{region 'Documentation'}
(*!
<summary>Advances a reconciled execution slot or dispatches one first-fitting Start; no owner lifecycle changes.</summary>
*)
{endregion}
METHOD PRIVATE ProcessSlot
IF (FResult = E_Result.Error) OR FExecutionFinished THEN
    RETURN;
END_IF;
IF IsSlotCompleted() THEN
    IF IsLastSlot(Slot := FCurrentSlot) THEN
        FExecutionFinished := TRUE;
    ELSE
        SelectNextSlot();
    END_IF;
    RETURN;
END_IF;
StartNextChild();
END_METHOD

{region 'Documentation'}
(*!
<summary>Publishes technical events through the configured framework publisher.</summary>
*)
{endregion}
METHOD PRIVATE PublishEvent
VAR_INPUT
    Event : ST_Event; //! Technical event value forwarded to the selected publisher; this helper performs no retry.
END_VAR
EventPublisher.PublishEvent(Event := Event);
END_METHOD

{region 'Documentation'}
(*!
<summary>Reads one initialized child at a validated occupied index; reports invalid bindings.</summary>
*)
{endregion}
METHOD PRIVATE ReadChild : I_Orchestratable //! Initialized child interface at Index; zero on invalid access or binding, with a technical Error latched.
VAR_INPUT
    Index : DINT; //! Original array index within the cached occupied child range.
END_VAR
VAR
    Child : I_Orchestratable;
END_VAR
ReadChild := 0;
IF (FCollection = 0) OR (Index < FFirstOccupiedIndex) OR (Index > FLastOccupiedIndex) THEN
    Error(Message := CONCAT('Invalid collection access at index ', DINT_TO_STRING(Index)));
    RETURN;
END_IF;

Child := FCollection.GetChild(Index := Index);
IF Child = 0 THEN
    Error(Message := CONCAT('Missing child at index ', DINT_TO_STRING(Index)));
    RETURN;
END_IF;
IF NOT Child.IsInitialized THEN
    Error(Message := CONCAT('Uninitialized child: ', Child.Name));
    RETURN;
END_IF;

ReadChild := Child;
END_METHOD

{region 'Documentation'}
(*!
<summary>Dispatches at most one capacity-admitted Reset per call; already ready children are skipped.</summary>
*)
{endregion}
METHOD PRIVATE ResetNextChild
VAR
    Child : I_Orchestratable;
    Index : DINT;
    ReservationResult : E_EventReservationResult;
END_VAR
WHILE UDINT_TO_LINT(FNextResetOffset) < (DINT_TO_LINT(FLastOccupiedIndex) - DINT_TO_LINT(FFirstOccupiedIndex) + 1) DO
    Index := LINT_TO_DINT(DINT_TO_LINT(FFirstOccupiedIndex) + UDINT_TO_LINT(FNextResetOffset));
    Child := ReadChild(Index := Index);
    IF Child = 0 THEN
        FNextResetOffset := FNextResetOffset + 1;
        RETURN;
    END_IF;
    IF (Child.State = E_State.Idle) AND Child.IsReady THEN
        FNextResetOffset := FNextResetOffset + 1;
        CONTINUE;
    END_IF;

    ReservationResult := Child.ReserveResetEvents();
    CASE ReservationResult OF
        E_EventReservationResult.Accepted:
            Child.RequestReset();
            FNextResetOffset := FNextResetOffset + 1;
        E_EventReservationResult.WaitingForCapacity:
            RETURN;
    ELSE
        Error(Message := CONCAT('Invalid child Reset reservation: ', Child.Name));
        FNextResetOffset := FNextResetOffset + 1;
    END_CASE;
    RETURN;
END_WHILE;
END_METHOD

{region 'Documentation'}
(*!
<summary>Neutral or held technical Error; task completion is reported separately.</summary>
*)
{endregion}
{attribute 'monitoring' := 'call'}
PROPERTY PUBLIC Result : E_Result //! Neutral or held technical Error; task completion is reported separately.
GET // PUBLIC
Result := FResult;
END_GET
END_PROPERTY

{region 'Documentation'}
(*!
<summary>Selects the first or next contiguous slot group; the caller owns advancement timing.</summary>
*)
{endregion}
METHOD PRIVATE SelectNextSlot : BOOL //! TRUE after selecting a valid contiguous slot group; FALSE indicates a technical Error.
VAR
    FirstIndex : LINT;
    Slot : UDINT;
    LastIndex : DINT;
    Index : LINT;
    Child : I_Orchestratable;
    ChildSlot : UINT;
END_VAR
SelectNextSlot := FALSE;
IF FCurrentSlot = 0 THEN
    FirstIndex := DINT_TO_LINT(FFirstOccupiedIndex);
    Slot := 1;
ELSE
    FirstIndex := DINT_TO_LINT(FSlotLastIndex) + 1;
    Slot := UINT_TO_UDINT(FCurrentSlot) + 1;
END_IF;

IF (FirstIndex < DINT_TO_LINT(FFirstOccupiedIndex)) OR (FirstIndex > DINT_TO_LINT(FLastOccupiedIndex))
    OR (Slot = 0) OR (UDINT_TO_LINT(Slot) > (DINT_TO_LINT(FLastOccupiedIndex) - DINT_TO_LINT(FFirstOccupiedIndex) + 1)) THEN
    Error(Message := 'Invalid child slot boundary.');
    RETURN;
END_IF;

LastIndex := LINT_TO_DINT(FirstIndex);
FOR Index := FirstIndex TO DINT_TO_LINT(FLastOccupiedIndex) DO
    Child := ReadChild(Index := LINT_TO_DINT(Index));
    IF Child = 0 THEN
        RETURN;
    END_IF;
    ChildSlot := Child.ExecutionSlot;
    IF UINT_TO_UDINT(ChildSlot) = Slot THEN
        LastIndex := LINT_TO_DINT(Index);
        CONTINUE;
    END_IF;
    IF (Index = FirstIndex) OR (UINT_TO_UDINT(ChildSlot) <> Slot + 1) THEN
        Error(Message := 'Child slots are not contiguous and ordered.');
        RETURN;
    END_IF;
    EXIT;
END_FOR;
FCurrentSlot := UDINT_TO_UINT(Slot);
FSlotFirstIndex := LINT_TO_DINT(FirstIndex);
FSlotLastIndex := LastIndex;
SelectNextSlot := TRUE;
END_METHOD

{region 'Documentation'}
(*!
<summary>Reserves and requests at most one first-fitting Child Start within the current slot.</summary>
*)
{endregion}
METHOD PRIVATE StartNextChild
VAR
    Index : LINT;
    Child : I_Orchestratable;
    ReservationResult : E_EventReservationResult;
END_VAR
FOR Index := DINT_TO_LINT(FSlotFirstIndex) TO DINT_TO_LINT(FSlotLastIndex) DO
    Child := ReadChild(Index := LINT_TO_DINT(Index));
    IF Child = 0 THEN
        RETURN;
    END_IF;
    IF Child.State <> E_State.Idle THEN
        CONTINUE;
    END_IF;

    ReservationResult := Child.ReserveExecutionEvents();
    CASE ReservationResult OF
        E_EventReservationResult.Accepted:
            Child.RequestStart();
            FPendingStartIndex := LINT_TO_DINT(Index);
            FHasPendingStart := TRUE;
            RETURN;
        E_EventReservationResult.WaitingForCapacity:
            CONTINUE;
    ELSE
        Error(Message := CONCAT('Invalid child execution reservation: ', Child.Name));
        RETURN;
    END_CASE;
END_FOR;
END_METHOD

{region 'Documentation'}
(*!
<summary>Prepares abort completion from stopped children; no requests, diagnostics or reservation changes.</summary>
*)
{endregion}
METHOD PRIVATE UpdateAbortCompletion
VAR
    Index : LINT;
    Child : I_Orchestratable;
END_VAR
FAbortFinished := FALSE;
IF FCollection = 0 THEN
    RETURN;
END_IF;
FOR Index := DINT_TO_LINT(FFirstOccupiedIndex) TO DINT_TO_LINT(FLastOccupiedIndex) DO
    Child := FCollection.GetChild(Index := LINT_TO_DINT(Index));
    IF Child = 0 THEN
        RETURN;
    END_IF;
    IF NOT Child.IsInitialized THEN
        RETURN;
    END_IF;
    IF NOT (((Child.State = E_State.Idle) AND Child.IsReady)
        OR ((Child.State = E_State.Completed) AND Child.IsComplete)) THEN
        RETURN;
    END_IF;
END_FOR;
FAbortFinished := TRUE;
END_METHOD

{region 'Documentation'}
(*!
<summary>Prepares start readiness without interpreting previous-run results or changing children.</summary>
*)
{endregion}
METHOD PRIVATE UpdateReadiness
VAR
    Index : LINT;
    Child : I_Orchestratable;
END_VAR
FChildrenReady := FALSE;
IF FCollection = 0 THEN
    RETURN;
END_IF;
FOR Index := DINT_TO_LINT(FFirstOccupiedIndex) TO DINT_TO_LINT(FLastOccupiedIndex) DO
    Child := FCollection.GetChild(Index := LINT_TO_DINT(Index));
    IF Child = 0 THEN
        RETURN;
    END_IF;
    IF NOT Child.IsInitialized THEN
        RETURN;
    END_IF;
    IF (Child.State <> E_State.Idle) OR NOT Child.IsReady THEN
        RETURN;
    END_IF;
END_FOR;
FChildrenReady := TRUE;
END_METHOD

{region 'Documentation'}
(*!
<summary>Prepares reset completion only after all dispatch attempts; failed terminal children count as finished.</summary>
*)
{endregion}
METHOD PRIVATE UpdateResetCompletion
VAR
    Index : LINT;
    Child : I_Orchestratable;
END_VAR
FResetFinished := FALSE;
IF FCollection = 0 THEN
    RETURN;
END_IF;
IF UDINT_TO_LINT(FNextResetOffset) < (DINT_TO_LINT(FLastOccupiedIndex) - DINT_TO_LINT(FFirstOccupiedIndex) + 1) THEN
    RETURN;
END_IF;
FOR Index := DINT_TO_LINT(FFirstOccupiedIndex) TO DINT_TO_LINT(FLastOccupiedIndex) DO
    Child := FCollection.GetChild(Index := LINT_TO_DINT(Index));
    IF Child = 0 THEN
        RETURN;
    END_IF;
    IF NOT Child.IsInitialized THEN
        RETURN;
    END_IF;
    IF NOT (((Child.State = E_State.Idle) AND Child.IsReady)
        OR ((Child.State = E_State.Completed) AND Child.IsComplete)) THEN
        RETURN;
    END_IF;
END_FOR;
FResetFinished := TRUE;
END_METHOD

END_FUNCTION_BLOCK

// ---- Framework/EventBuffer/POU/FrameworkEvents/CreateFrameworkEvent.TcPOU
{region 'Documentation'}
(*!
<summary>Constructs a framework diagnostic event without publishing it.</summary>
<description>
Name and Message are ASCII text limited to the declared event capacities.
</description>
*)
{endregion}
FUNCTION CreateFrameworkEvent : ST_Event //! Constructed event value; not published. The publisher assigns SequenceId and Timestamp.
VAR_INPUT
    Name : STRING(GVL_Constants.NameLength); //! Hierarchical owner name used to identify events; must satisfy the naming contract.
    ResourceName : STRING(GVL_Constants.ResourceNameLength) := ''; //! Optional resource context for diagnostics; empty by default.
    State : E_State; //! Owner lifecycle state recorded in the event.
    Severity : E_EventSeverity; //! Logging severity for the diagnostic; independent of the test result.
    Message : STRING(GVL_Constants.MessageLength); //! Diagnostic text copied into the event within MessageLength.
END_VAR

CreateFrameworkEvent.SequenceId := 0;
CreateFrameworkEvent.Timestamp := 0;
CreateFrameworkEvent.OwnerScope := E_OwnerScope.Framework;
CreateFrameworkEvent.EventType := E_EventType.Framework;
CreateFrameworkEvent.Severity := Severity;
CreateFrameworkEvent.Name := Name;
CreateFrameworkEvent.ResourceName := ResourceName;
CreateFrameworkEvent.State := State;
CreateFrameworkEvent.Result := E_Result.NotEvaluated;
CreateFrameworkEvent.Message := Message;

END_FUNCTION

// ---- Framework/Common/POU/Stopwatch.TcPOU
{region 'Documentation'}
(*!
<summary>Internal method-driven duration measurement; no FB-body call is required. Start/Update/Stop use the current task&#x27;s scheduled timestamp. Reset clears the measurement. ElapsedTicks retains 100 ns resolution; ElapsedTime is the saturated millisecond projection.</summary>
<description>
Start replaces the previous interval. Update samples only while running and valid; Stop performs one final Update. A backward task timestamp latches invalid until Start or Reset. Property reads return held values rather than sampling the clock. ElapsedLTime is a direct conversion, without the saturation applied to ElapsedTime.


The source is the current task's scheduled timestamp, so this measures elapsed task time rather than execution cost between operations within the same task cycle. Check IsValid before using a refreshed value; a backward observation leaves the last valid duration held and does not repair itself on later Update calls.
</description>
*)
{endregion}
FUNCTION_BLOCK INTERNAL Stopwatch
VAR
    FRunning : BOOL;
    FIsValid : BOOL := TRUE;
    FStartTicks : ULINT;
    FPreviousTicks : ULINT;
    FElapsedTicks : ULINT;
END_VAR

{region 'Documentation'}
(*!
<summary>Nanosecond projection of the last updated 100 ns duration; reading does not refresh the measurement.</summary>
*)
{endregion}
{attribute 'monitoring' := 'call'}
PROPERTY PUBLIC ElapsedLTime : LTIME //! Held duration converted to LTIME nanoseconds; no refresh on read.
GET // PUBLIC
ElapsedLTime := ULINT_TO_LTIME(FElapsedTicks * 100);
END_GET
END_PROPERTY

{region 'Documentation'}
(*!
<summary>Elapsed duration in 100 ns ticks from the latest Start, Update or Stop; reading does not sample the clock.</summary>
*)
{endregion}
{attribute 'monitoring' := 'call'}
PROPERTY PUBLIC ElapsedTicks : ULINT //! Held elapsed duration in 100 ns ticks; no refresh on read.
GET // PUBLIC
ElapsedTicks := FElapsedTicks;
END_GET
END_PROPERTY

{region 'Documentation'}
(*!
<summary>Millisecond projection of the last updated duration, saturated at TIME's maximum value; reading does not refresh it.</summary>
*)
{endregion}
{attribute 'monitoring' := 'call'}
PROPERTY PUBLIC ElapsedTime : TIME //! Held duration in milliseconds, saturated at TIME's maximum; no refresh on read.
GET // PUBLIC
VAR CONSTANT
	MaxTime: ULINT := 42949672950000;
END_VAR
ElapsedTime := ULINT_TO_TIME(MIN(FElapsedTicks, MaxTime) / 10000);
END_GET
END_PROPERTY

{region 'Documentation'}
(*!
<summary>Report whether a backward clock observation has invalidated the measurement; Start or Reset restores validity.</summary>
*)
{endregion}
{attribute 'monitoring' := 'call'}
PROPERTY PUBLIC IsValid : BOOL //! FALSE after Update observes backward time; latched until Start or Reset.
GET // PUBLIC
IsValid := FIsValid;
END_GET
END_PROPERTY

{region 'Documentation'}
(*!
<summary>Clears the held measurement without starting a new interval.</summary>
*)
{endregion}
METHOD PUBLIC Reset
FRunning := FALSE;
FIsValid := TRUE;
FStartTicks := 0;
FPreviousTicks := 0;
FElapsedTicks := 0;
END_METHOD

{region 'Documentation'}
(*!
<summary>Starts a new measurement, replacing the previous value.</summary>
*)
{endregion}
METHOD PUBLIC Start
FStartTicks := Tc2_System.F_GetTaskTime();
FPreviousTicks := FStartTicks;
FElapsedTicks := 0;
FIsValid := TRUE;
FRunning := TRUE;
END_METHOD

{region 'Documentation'}
(*!
<summary>Captures the final duration and holds it until the next Start or Reset.</summary>
<description>
If the final Update detects backward time, IsValid becomes FALSE and the last valid elapsed value remains held. Stop still ends the interval. Repeated Stop calls do not sample again while stopped.
</description>
*)
{endregion}
METHOD PUBLIC Stop
Update();
FRunning := FALSE;
END_METHOD

{region 'Documentation'}
(*!
<summary>Refreshes elapsed time. A backwards clock latches invalid until Start or Reset.</summary>
*)
{endregion}
METHOD PUBLIC Update
VAR
    Ticks : ULINT;
END_VAR
IF NOT FRunning OR NOT FIsValid THEN
    RETURN;
END_IF;
Ticks := Tc2_System.F_GetTaskTime();
IF Ticks < FPreviousTicks THEN
    FIsValid := FALSE;
    RETURN;
END_IF;

FElapsedTicks := Ticks - FStartTicks;
FPreviousTicks := Ticks;
END_METHOD

END_FUNCTION_BLOCK

// ---- Framework/Common/POU/ResultAggregator.TcPOU
{region 'Documentation'}
(*!
<summary>Incrementally collect results through methods; no cyclic FB call is required. Reset starts an empty collection; Add methods always contribute. Each contribution counts once; the owner limits each collection to the UINT range.</summary>
<description>
Use Reset before each new collection and contribute each intended provider/result exactly once. AddProvider reads immediately and retains no interface. Error has highest precedence but does not stop later counter updates. TotalCount includes NotEvaluated and Abort contributions, so PassedCount, FailedCount and ErrorCount do not necessarily sum to TotalCount. The caller keeps a collection within 65535 contributions; counters are not saturating. This object emits no events and does not execute providers.
</description>
*)
{endregion}
FUNCTION_BLOCK ResultAggregator IMPLEMENTS I_ResultAggregator
VAR
    FResult : E_Result := E_Result.NotEvaluated;
    FTotalCount : UINT;
    FPassedCount : UINT;
    FFailedCount : UINT;
    FErrorCount : UINT;
END_VAR

{region 'Documentation'}
(*!
<summary>Adds one provider result; a null provider contributes one Error. Reads the result immediately; no reference is retained.</summary>
*)
{endregion}
METHOD PUBLIC AddProvider
VAR_INPUT
    Provider : I_ResultProvider; //! Result provider read immediately; zero contributes Error. No reference is retained.
END_VAR
IF Provider = 0 THEN
    AddResult(Result := E_Result.Error);
    RETURN;
END_IF;
AddResult(Result := Provider.Result);
END_METHOD

{region 'Documentation'}
(*!
<summary>Counts one contribution and combines Error &gt; Abort &gt; Failed &gt; Passed &gt; NotEvaluated.</summary>
*)
{endregion}
METHOD PUBLIC AddResult
VAR_INPUT
    Result : E_Result; //! Evaluation result to count as one contribution; severity is Error > Abort > Failed > Passed > NotEvaluated.
END_VAR
FTotalCount := FTotalCount + 1;
CASE Result OF
    E_Result.Passed:
        FPassedCount := FPassedCount + 1;
    E_Result.Failed:
        FFailedCount := FFailedCount + 1;
    E_Result.Error:
        FErrorCount := FErrorCount + 1;
END_CASE;

IF FResult = E_Result.Error THEN
    RETURN;
END_IF;

CASE Result OF
    E_Result.NotEvaluated:
        RETURN;
    E_Result.Passed:
        IF FResult = E_Result.NotEvaluated THEN
            FResult := Result;
        END_IF;
    E_Result.Failed:
        IF FResult <> E_Result.Abort THEN
            FResult := Result;
        END_IF;
    E_Result.Abort, E_Result.Error:
        FResult := Result;
END_CASE;
END_METHOD

{region 'Documentation'}
(*!
<summary>Number of accepted Error contributions.</summary>
*)
{endregion}
{attribute 'monitoring' := 'call'}
PROPERTY PUBLIC ErrorCount : UINT //! Number of accepted Error contributions.
GET // PUBLIC
ErrorCount := FErrorCount;
END_GET
END_PROPERTY

{region 'Documentation'}
(*!
<summary>Number of accepted Failed contributions.</summary>
*)
{endregion}
{attribute 'monitoring' := 'call'}
PROPERTY PUBLIC FailedCount : UINT //! Number of accepted Failed contributions.
GET // PUBLIC
FailedCount := FFailedCount;
END_GET
END_PROPERTY

{region 'Documentation'}
(*!
<summary>Number of accepted Passed contributions.</summary>
*)
{endregion}
{attribute 'monitoring' := 'call'}
PROPERTY PUBLIC PassedCount : UINT //! Number of accepted Passed contributions.
GET // PUBLIC
PassedCount := FPassedCount;
END_GET
END_PROPERTY

{region 'Documentation'}
(*!
<summary>Starts an empty collection by clearing result and counters immediately.</summary>
*)
{endregion}
METHOD PUBLIC Reset
FResult := E_Result.NotEvaluated;
FTotalCount := 0;
FPassedCount := 0;
FFailedCount := 0;
FErrorCount := 0;
END_METHOD

{region 'Documentation'}
(*!
<summary>Current aggregate; an empty collection is NotEvaluated.</summary>
*)
{endregion}
{attribute 'monitoring' := 'call'}
PROPERTY PUBLIC Result : E_Result //! Current aggregate; an empty collection is NotEvaluated.
GET // PUBLIC
Result := FResult;
END_GET
END_PROPERTY

{region 'Documentation'}
(*!
<summary>Number of accepted contributions, including NotEvaluated and Abort.</summary>
*)
{endregion}
{attribute 'monitoring' := 'call'}
PROPERTY PUBLIC TotalCount : UINT //! Number of accepted contributions, including NotEvaluated and Abort.
GET // PUBLIC
TotalCount := FTotalCount;
END_GET
END_PROPERTY

END_FUNCTION_BLOCK

// ---- Framework/EventBuffer/POU/FrameworkEvents/CreateInvalidStateTransitionEvent.TcPOU
{region 'Documentation'}
(*!
<summary>Constructs a Framework Error diagnostic for a rejected transition without publishing it.</summary>
<description>
State records StateOld; Message includes StateOld and the rejected StateNew. No transition is performed.
</description>
*)
{endregion}
FUNCTION CreateInvalidStateTransitionEvent : ST_Event //! Constructed event value; not published. The publisher assigns SequenceId and Timestamp.
VAR_INPUT
    OwnerScope : E_OwnerScope; //! Semantic owner category recorded in the event.
    Name : STRING(GVL_Constants.NameLength); //! Hierarchical owner name used to identify events; must satisfy the naming contract.
    ResourceName : STRING(GVL_Constants.ResourceNameLength) := ''; //! Optional resource context for diagnostics; empty by default.
    StateOld : E_State; //! Owner state before the reported or rejected transition.
    StateNew : E_State; //! Rejected destination included in Message; the structured event State remains StateOld.
END_VAR
VAR
    Message : STRING(GVL_Constants.MessageLength);
END_VAR

Message := CONCAT(STR1 := 'Invalid State transition requested ', STR2 := INT_TO_STRING(TO_INT(StateOld)));
Message := CONCAT(STR1 := Message, STR2 := ' -> ');
Message := CONCAT(STR1 := Message, STR2 := INT_TO_STRING(TO_INT(StateNew)));

CreateInvalidStateTransitionEvent.SequenceId := 0;
CreateInvalidStateTransitionEvent.Timestamp := 0;
CreateInvalidStateTransitionEvent.OwnerScope := OwnerScope;
CreateInvalidStateTransitionEvent.EventType := E_EventType.Framework;
CreateInvalidStateTransitionEvent.Severity := E_EventSeverity.Error;
CreateInvalidStateTransitionEvent.Name := Name;
CreateInvalidStateTransitionEvent.ResourceName := ResourceName;
CreateInvalidStateTransitionEvent.State := StateOld;
CreateInvalidStateTransitionEvent.Result := E_Result.NotEvaluated;
CreateInvalidStateTransitionEvent.Message := Message;

END_FUNCTION

// ---- Framework/EventBuffer/POU/FrameworkEvents/CreateResetWarningEvent.TcPOU
{region 'Documentation'}
(*!
<summary>Constructs a Framework Warning diagnostic for Reset interrupting an active owner lifecycle.</summary>
<description>
State identifies the interrupted state. The function neither publishes the event nor performs Reset.
</description>
*)
{endregion}
FUNCTION CreateResetWarningEvent : ST_Event //! Constructed event value; not published. The publisher assigns SequenceId and Timestamp.
VAR_INPUT
    OwnerScope : E_OwnerScope; //! Semantic owner category recorded in the event.
	Name : STRING(GVL_Constants.NameLength); //! Hierarchical owner name used to identify events; must satisfy the naming contract.
    ResourceName : STRING(GVL_Constants.ResourceNameLength) := ''; //! Optional resource context for diagnostics; empty by default.
    State : E_State; //! Owner lifecycle state recorded in the event.
END_VAR
VAR
    Message : STRING(GVL_Constants.MessageLength);
END_VAR

CASE OwnerScope OF
	E_OwnerScope.Preparation: Message := 'Reset interrupts an active Preparation lifecycle.';
	E_OwnerScope.TestCase: Message := 'Reset interrupts an active Test Case lifecycle.';
	E_OwnerScope.TestSuite: Message := 'Reset interrupts an active Test Suite lifecycle.';
	E_OwnerScope.RunControl: Message := 'Reset interrupts an active Unit Test lifecycle.';
	ELSE Message := 'Reset interrupts an active owner lifecycle.';
END_CASE


CreateResetWarningEvent.SequenceId := 0;
CreateResetWarningEvent.Timestamp := 0;
CreateResetWarningEvent.OwnerScope := OwnerScope;
CreateResetWarningEvent.EventType := E_EventType.Framework;
CreateResetWarningEvent.Severity := E_EventSeverity.Warning;
CreateResetWarningEvent.Name := Name;
CreateResetWarningEvent.ResourceName := ResourceName;
CreateResetWarningEvent.State := State;
CreateResetWarningEvent.Result := E_Result.NOTEVALUATED;
CreateResetWarningEvent.Message := Message;

END_FUNCTION

// ---- Framework/EventBuffer/POU/StateTransitionEvents/CreateStateTransitionEvent.TcPOU
{region 'Documentation'}
(*!
<summary>Constructs an owner state-transition event without publishing it.</summary>
<description>
The caller supplies valid ASCII owner context; the structured state is StateNew.
</description>
*)
{endregion}
FUNCTION CreateStateTransitionEvent : ST_Event //! Constructed event value; not published. The publisher assigns SequenceId and Timestamp.
VAR_INPUT
    OwnerScope : E_OwnerScope; //! Semantic owner category recorded in the event.
    Name : STRING(GVL_Constants.NameLength); //! Hierarchical owner name used to identify events; must satisfy the naming contract.
    ResourceName : STRING(GVL_Constants.ResourceNameLength) := ''; //! Optional resource context for diagnostics; empty by default.
    StateOld : E_State; //! Owner state before the reported or rejected transition.
    StateNew : E_State; //! Requested destination state recorded in the event; this function does not perform the transition.
END_VAR

CreateStateTransitionEvent.SequenceId := 0;
CreateStateTransitionEvent.Timestamp := 0;
CreateStateTransitionEvent.OwnerScope := OwnerScope;
CreateStateTransitionEvent.EventType := E_EventType.StateTransition;
CreateStateTransitionEvent.Severity := E_EventSeverity.Info;
CreateStateTransitionEvent.Name := Name;
CreateStateTransitionEvent.ResourceName := ResourceName;
CreateStateTransitionEvent.State := StateNew;
CreateStateTransitionEvent.Result := E_Result.NotEvaluated;
CreateStateTransitionEvent.Message := CONCAT(STR1 := 'State transition ',
    STR2 := INT_TO_STRING(TO_INT(StateOld)));
CreateStateTransitionEvent.Message := CONCAT(STR1 := CreateStateTransitionEvent.Message,
    STR2 := ' -> ');
CreateStateTransitionEvent.Message := CONCAT(STR1 := CreateStateTransitionEvent.Message,
    STR2 := INT_TO_STRING(TO_INT(StateNew)));

END_FUNCTION

// ---- Framework/RunControl/POU/RunControlConfigurationBuilder.TcPOU
{region 'Documentation'}
(*!
<summary>Setup-only configuration: Initialize through Finalize requires stable array/child storage.</summary>
<description>
No FB body call is required. Finalize discards the temporary array pointer on either outcome.
At most 65535 children can be registered; Initialize clears the complete array after validating mode and capacity.


The returned configuration describes the owner's actual array; Finalize does not copy child storage or make it immutable. Keep that array, child instances and assigned slots stable for the complete execution lifetime. Do not retain a temporary builder passed to Configure. Setup clears array capacity and scans/shifts registered entries; it is configuration work, not cyclic scheduling.
</description>
*)
{endregion}
FUNCTION_BLOCK RunControlConfigurationBuilder
VAR
    FInitialized : BOOL;
    FEntries : POINTER TO I_TestSuite;
    FFinalized : BOOL;
    FRegistrationError : BOOL;
    FConfiguration : ST_TestSuiteCollectionConfig;
END_VAR

VAR CONSTANT
    MaxCount : UINT := 65535;
END_VAR

{region 'Documentation'}
(*!
<summary>Number of registered entries, contiguous from FirstIndex.</summary>
*)
{endregion}
{attribute 'monitoring' := 'call'}
PROPERTY PUBLIC Count : UINT //! Number of registered entries, contiguous from FirstIndex.
GET // PUBLIC
Count := FConfiguration.Count;
END_GET
END_PROPERTY

{region 'Documentation'}
(*!
<summary>Finalizes validation and releases the array binding; repeated calls return the same configuration.</summary>
<description>
An empty collection or any latched registration error is invalid. Serial slots must follow registration order; Parallel uses slot one; ParallelSlots must form consecutive positive groups starting at one. The temporary pointer is discarded on every first finalization outcome. Finalization validates slots and bindings, not child initialization; Run Control performs those later checks.
</description>
*)
{endregion}
METHOD PUBLIC Finalize : ST_TestSuiteCollectionConfig //! Finalized bounds, count and mode; IsValid determines whether the configuration can be used.
VAR
    Offset : DINT;
    PreviousSlot : UDINT;
    Slot : UDINT;
    Child : I_TestSuite;
END_VAR
IF FFinalized THEN
    Finalize := FConfiguration;
    RETURN;
END_IF;

IF NOT FInitialized OR FRegistrationError OR (FEntries = 0) OR (FConfiguration.Count = 0) THEN
    FConfiguration.IsValid := FALSE;
    FEntries := 0;
    FFinalized := TRUE;
    Finalize := FConfiguration;
    RETURN;
END_IF;

PreviousSlot := 0;
FOR Offset := 0 TO UINT_TO_DINT(FConfiguration.Count) - 1 DO
    Child := FEntries[Offset];
    IF Child = 0 THEN
        FRegistrationError := TRUE;
        EXIT;
    END_IF;
    Slot := UINT_TO_UDINT(Child.ExecutionSlot);
    IF (Slot = 0) OR (Slot < PreviousSlot) OR (Slot > PreviousSlot + 1)
        OR ((FConfiguration.Mode = E_OrchestrationMode.Serial) AND (Slot <> DINT_TO_UDINT(Offset) + 1))
        OR ((FConfiguration.Mode = E_OrchestrationMode.Parallel) AND (Slot <> 1)) THEN
        FRegistrationError := TRUE;
        EXIT;
    END_IF;
    PreviousSlot := Slot;
END_FOR;

FConfiguration.IsValid := NOT FRegistrationError;
FEntries := 0;
FFinalized := TRUE;
Finalize := FConfiguration;
END_METHOD

{region 'Documentation'}
(*!
<summary>Actual lower bound of the supplied array.</summary>
*)
{endregion}
{attribute 'monitoring' := 'call'}
PROPERTY PUBLIC FirstIndex : DINT //! Actual lower bound of the supplied array.
GET // PUBLIC
FirstIndex := FConfiguration.FirstIndex;
END_GET
END_PROPERTY

{region 'Documentation'}
(*!
<summary>Starts a new build and clears the supplied array; bounds and mode remain fixed until Finalize.</summary>
<description>
A valid mode and a positive array capacity are checked before the array is cleared; rejected prerequisites leave its entries untouched. Registration starts at the actual lower bound and occupies a contiguous prefix. A new Initialize starts a fresh build after previous success or failure. The registration count is capped at 65535 even if physical capacity is larger.
</description>
*)
{endregion}
METHOD PUBLIC Initialize
VAR_INPUT
    Mode : E_OrchestrationMode; //! Scheduling strategy fixed for this build; Register is for Serial/Parallel, RegisterWithSlot for ParallelSlots.
END_VAR
VAR_IN_OUT
    TestSuites : ARRAY[*] OF I_TestSuite; //! Owner-held array cleared and filled by the builder; storage must stay fixed through Finalize and registered children must outlive execution.
END_VAR
VAR
    Index : LINT;
    Capacity : LINT;
END_VAR
FInitialized := FALSE;
FEntries := 0;
FFinalized := FALSE;
FRegistrationError := FALSE;
FConfiguration.IsValid := FALSE;
FConfiguration.Count := 0;
FConfiguration.FirstIndex := LOWER_BOUND(TestSuites, 1);
FConfiguration.LastIndex := UPPER_BOUND(TestSuites, 1);
FConfiguration.Mode := Mode;

IF (Mode <> E_OrchestrationMode.Serial)
    AND (Mode <> E_OrchestrationMode.Parallel)
    AND (Mode <> E_OrchestrationMode.ParallelSlots) THEN
    FRegistrationError := TRUE;
    RETURN;
END_IF;

Capacity := DINT_TO_LINT(FConfiguration.LastIndex) - DINT_TO_LINT(FConfiguration.FirstIndex) + 1;
IF Capacity <= 0 THEN
    FRegistrationError := TRUE;
    RETURN;
END_IF;

FOR Index := DINT_TO_LINT(FConfiguration.FirstIndex) TO DINT_TO_LINT(FConfiguration.LastIndex) DO
    TestSuites[LINT_TO_DINT(Index)] := 0;
END_FOR;
FEntries := ADR(TestSuites[FConfiguration.FirstIndex]);
FInitialized := TRUE;
END_METHOD

{region 'Documentation'}
(*!
<summary>Validates before mutation, inserts the child and sets its effective slot.</summary>
*)
{endregion}
METHOD PRIVATE Insert : BOOL //! TRUE after insertion and slot assignment; FALSE latches a registration error without adding an entry.
VAR_INPUT
    TestSuite : I_TestSuite; //! Unique nonzero child to insert; the instance must outlive the finalized owner collection.
    ExecutionSlot : UINT; //! Positive effective slot; stable sorted insertion preserves registration order within equal slots.
END_VAR
VAR
    Offset : DINT;
    InsertOffset : DINT;
    Child : I_TestSuite;
END_VAR
Insert := FALSE;
IF NOT FInitialized OR FRegistrationError OR (FEntries = 0) OR (TestSuite = 0) OR (ExecutionSlot = 0) THEN
    FRegistrationError := TRUE;
    RETURN;
END_IF;
IF (FConfiguration.Count = MaxCount)
    OR (UINT_TO_LINT(FConfiguration.Count) >= DINT_TO_LINT(FConfiguration.LastIndex) - DINT_TO_LINT(FConfiguration.FirstIndex) + 1) THEN
    FRegistrationError := TRUE;
    RETURN;
END_IF;

InsertOffset := UINT_TO_DINT(FConfiguration.Count);
FOR Offset := 0 TO UINT_TO_DINT(FConfiguration.Count) - 1 DO
    Child := FEntries[Offset];
    IF (Child = 0) OR (Child = TestSuite) THEN
        FRegistrationError := TRUE;
        RETURN;
    END_IF;
    IF (InsertOffset = UINT_TO_DINT(FConfiguration.Count)) AND (Child.ExecutionSlot > ExecutionSlot) THEN
        InsertOffset := Offset;
    END_IF;
END_FOR;
IF FEntries[FConfiguration.Count] <> 0 THEN
    FRegistrationError := TRUE;
    RETURN;
END_IF;

TestSuite.ExecutionSlot := ExecutionSlot;
FOR Offset := UINT_TO_DINT(FConfiguration.Count) TO InsertOffset + 1 BY -1 DO
    FEntries[Offset] := FEntries[Offset - 1];
END_FOR;
FEntries[InsertOffset] := TestSuite;
FConfiguration.Count := FConfiguration.Count + 1;
Insert := TRUE;
END_METHOD

{region 'Documentation'}
(*!
<summary>Finalize has completed, independently of validation success.</summary>
*)
{endregion}
{attribute 'monitoring' := 'call'}
PROPERTY PUBLIC IsFinalized : BOOL //! Finalize has completed, independently of validation success.
GET // PUBLIC
IsFinalized := FFinalized;
END_GET
END_PROPERTY

{region 'Documentation'}
(*!
<summary>Finalization succeeded; FALSE before Finalize.</summary>
*)
{endregion}
{attribute 'monitoring' := 'call'}
PROPERTY PUBLIC IsValid : BOOL //! Finalization succeeded; FALSE before Finalize.
GET // PUBLIC
IsValid := FConfiguration.IsValid;
END_GET
END_PROPERTY

{region 'Documentation'}
(*!
<summary>Actual upper bound, including unused capacity.</summary>
*)
{endregion}
{attribute 'monitoring' := 'call'}
PROPERTY PUBLIC LastIndex : DINT //! Actual upper bound, including unused capacity.
GET // PUBLIC
LastIndex := FConfiguration.LastIndex;
END_GET
END_PROPERTY

{region 'Documentation'}
(*!
<summary>Mode selected by Initialize.</summary>
*)
{endregion}
{attribute 'monitoring' := 'call'}
PROPERTY PUBLIC Mode : E_OrchestrationMode //! Mode selected by Initialize.
GET // PUBLIC
Mode := FConfiguration.Mode;
END_GET
END_PROPERTY

{region 'Documentation'}
(*!
<summary>Appends a unique child in Serial or Parallel mode and assigns its effective slot.</summary>
<description>
Serial assigns increasing slots and Parallel assigns slot one. Rejection before finalization latches a build error, making Finalize invalid until another Initialize. After Finalize this method returns FALSE without altering the frozen configuration or adding a new error.
</description>
*)
{endregion}
METHOD PUBLIC Register : BOOL //! TRUE when the child was registered; FALSE adds no entry; pre-finalization rejection latches a build error.
VAR_INPUT
    TestSuite : I_TestSuite; //! Nonzero child interface to register once; its instance must outlive the registered collection.
END_VAR
VAR
    Slot : UINT;
END_VAR
Register := FALSE;
IF FFinalized THEN
    RETURN;
END_IF;
IF (FConfiguration.Mode <> E_OrchestrationMode.Serial)
    AND (FConfiguration.Mode <> E_OrchestrationMode.Parallel) THEN
    FRegistrationError := TRUE;
    RETURN;
END_IF;

Slot := 1;
IF FConfiguration.Mode = E_OrchestrationMode.Serial THEN
    IF FConfiguration.Count = MaxCount THEN
        FRegistrationError := TRUE;
        RETURN;
    END_IF;
    Slot := FConfiguration.Count + 1;
END_IF;
Register := Insert(TestSuite := TestSuite,
    ExecutionSlot := Slot);
END_METHOD

{region 'Documentation'}
(*!
<summary>Registers a unique child in ParallelSlots mode, stably inserting by positive slot.</summary>
<description>
Available only in ParallelSlots mode. Slots must be positive; stable insertion sorts the array by slot. Finalize additionally rejects gaps or a first slot other than one. Rejection before finalization latches a build error; calls after Finalize return FALSE without changing its frozen outcome.
</description>
*)
{endregion}
METHOD PUBLIC RegisterWithSlot : BOOL //! TRUE when the child was registered; FALSE adds no entry; pre-finalization rejection latches a build error.
VAR_INPUT
    TestSuite : I_TestSuite; //! Nonzero child interface to register once; its instance must outlive the registered collection.
    ExecutionSlot : UINT; //! Positive slot number for ParallelSlots registration; children sharing a slot may overlap, with at most one new Start admitted per helper call.
END_VAR
RegisterWithSlot := FALSE;
IF FFinalized THEN
    RETURN;
END_IF;
IF FConfiguration.Mode <> E_OrchestrationMode.ParallelSlots THEN
    FRegistrationError := TRUE;
    RETURN;
END_IF;
RegisterWithSlot := Insert(TestSuite := TestSuite,
    ExecutionSlot := ExecutionSlot);
END_METHOD

END_FUNCTION_BLOCK

// ---- Framework/EventBuffer/POU/ResultEvents/CreateResultEvent.TcPOU
{region 'Documentation'}
(*!
<summary>Constructs a result event without evaluating or publishing it.</summary>
<description>
The caller supplies the complete ASCII name, resource context and finding message.
</description>
*)
{endregion}
FUNCTION CreateResultEvent : ST_Event //! Constructed event value; not published. The publisher assigns SequenceId and Timestamp.
VAR_INPUT
    OwnerScope : E_OwnerScope; //! Semantic owner category recorded in the event.
    Name : STRING(GVL_Constants.NameLength); //! Hierarchical owner name used to identify events; must satisfy the naming contract.
    ResourceName : STRING(GVL_Constants.ResourceNameLength) := ''; //! Optional resource context for diagnostics; empty by default.
    State : E_State; //! Owner lifecycle state recorded in the event.
    Result : E_Result; //! Evaluation result to include or classify; its numeric value is not severity order.
    Message : STRING(GVL_Constants.MessageLength); //! Diagnostic text copied into the event within MessageLength.
END_VAR

CreateResultEvent.SequenceId := 0;
CreateResultEvent.Timestamp := 0;
CreateResultEvent.OwnerScope := OwnerScope;
CreateResultEvent.EventType := E_EventType.Result;
CreateResultEvent.Severity := SelectResultSeverity(Result := Result);
CreateResultEvent.Name := Name;
CreateResultEvent.ResourceName := ResourceName;
CreateResultEvent.State := State;
CreateResultEvent.Result := Result;
CreateResultEvent.Message := Message;

END_FUNCTION

// ---- Framework/EventBuffer/POU/Utilities/SelectResultSeverity.TcPOU
{region 'Documentation'}
(*!
<summary>Maps an evaluation result to logging severity, not result severity.</summary>
<description>
Passed and Failed map to Info; NotEvaluated and Abort map to Warning. Error and all other values map to Error. Logging severity is independent of the result aggregation order.
</description>
*)
{endregion}
FUNCTION INTERNAL SelectResultSeverity : E_EventSeverity //! Logging severity corresponding to Result.
VAR_INPUT
    Result : E_Result; //! Evaluation result to include or classify; its numeric value is not severity order.
END_VAR

CASE Result OF
    E_Result.NotEvaluated,
    E_Result.Abort:
        SelectResultSeverity := E_EventSeverity.Warning;
    E_Result.Passed,
    E_Result.Failed:
        SelectResultSeverity := E_EventSeverity.Info;
ELSE
    SelectResultSeverity := E_EventSeverity.Error;
END_CASE;

END_FUNCTION

// ---- Framework/EventBuffer/POU/AggregationEvents/CreateRunAggregationEvent.TcPOU
{region 'Documentation'}
(*!
<summary>Constructs a Run aggregation event from an already aggregated status snapshot.</summary>
<description>
Runtime is rendered as unsigned milliseconds; the caller owns publication.


Compact JSON fields are total, inactive, idle, running, completed, passed, failed, error, runtime and lostEvents. Counts and runtime are unsigned decimal numbers. This formats the supplied snapshot without validating completion or recomputing aggregation; the owner controls finalization order and publication.
</description>
*)
{endregion}
FUNCTION CreateRunAggregationEvent : ST_Event //! Constructed event value; not published. The publisher assigns SequenceId and Timestamp.
VAR_INPUT
    Name : STRING(GVL_Constants.NameLength); //! Hierarchical owner name used to identify events; must satisfy the naming contract.
    Status : ST_RunControlStatus; //! Already aggregated owner status snapshot; the function formats it without observing children.
    LostEventCount : UINT; //! Publisher's cumulative lost-event count included in the Run aggregation.
END_VAR
VAR
    RuntimeMilliseconds : UDINT;
END_VAR

RuntimeMilliseconds := TIME_TO_UDINT(Status.Runtime);

CreateRunAggregationEvent.SequenceId := 0;
CreateRunAggregationEvent.Timestamp := 0;
CreateRunAggregationEvent.OwnerScope := E_OwnerScope.RunControl;
CreateRunAggregationEvent.EventType := E_EventType.Aggregation;
CreateRunAggregationEvent.Severity := SelectResultSeverity(Result := Status.Execution.Result);
CreateRunAggregationEvent.Name := Name;
CreateRunAggregationEvent.ResourceName := '';
CreateRunAggregationEvent.State := Status.Execution.State;
CreateRunAggregationEvent.Result := Status.Execution.Result;

CreateRunAggregationEvent.Message := CONCAT(STR1 := '{"total":',
    STR2 := UINT_TO_STRING(Status.SuiteCountTotal));
CreateRunAggregationEvent.Message := CONCAT(STR1 := CreateRunAggregationEvent.Message,
    STR2 := ',"inactive":');
CreateRunAggregationEvent.Message := CONCAT(STR1 := CreateRunAggregationEvent.Message,
    STR2 := UINT_TO_STRING(Status.SuiteCountInactive));
CreateRunAggregationEvent.Message := CONCAT(STR1 := CreateRunAggregationEvent.Message,
    STR2 := ',"idle":');
CreateRunAggregationEvent.Message := CONCAT(STR1 := CreateRunAggregationEvent.Message,
    STR2 := UINT_TO_STRING(Status.SuiteCountIdle));
CreateRunAggregationEvent.Message := CONCAT(STR1 := CreateRunAggregationEvent.Message,
    STR2 := ',"running":');
CreateRunAggregationEvent.Message := CONCAT(STR1 := CreateRunAggregationEvent.Message,
    STR2 := UINT_TO_STRING(Status.SuiteCountRunning));
CreateRunAggregationEvent.Message := CONCAT(STR1 := CreateRunAggregationEvent.Message,
    STR2 := ',"completed":');
CreateRunAggregationEvent.Message := CONCAT(STR1 := CreateRunAggregationEvent.Message,
    STR2 := UINT_TO_STRING(Status.SuiteCountCompleted));
CreateRunAggregationEvent.Message := CONCAT(STR1 := CreateRunAggregationEvent.Message,
    STR2 := ',"passed":');
CreateRunAggregationEvent.Message := CONCAT(STR1 := CreateRunAggregationEvent.Message,
    STR2 := UINT_TO_STRING(Status.SuiteCountPassed));
CreateRunAggregationEvent.Message := CONCAT(STR1 := CreateRunAggregationEvent.Message,
    STR2 := ',"failed":');
CreateRunAggregationEvent.Message := CONCAT(STR1 := CreateRunAggregationEvent.Message,
    STR2 := UINT_TO_STRING(Status.SuiteCountFailed));
CreateRunAggregationEvent.Message := CONCAT(STR1 := CreateRunAggregationEvent.Message,
    STR2 := ',"error":');
CreateRunAggregationEvent.Message := CONCAT(STR1 := CreateRunAggregationEvent.Message,
    STR2 := UINT_TO_STRING(Status.SuiteCountError));
CreateRunAggregationEvent.Message := CONCAT(STR1 := CreateRunAggregationEvent.Message,
    STR2 := ',"runtime":');
CreateRunAggregationEvent.Message := CONCAT(STR1 := CreateRunAggregationEvent.Message,
    STR2 := UDINT_TO_STRING(RuntimeMilliseconds));
CreateRunAggregationEvent.Message := CONCAT(STR1 := CreateRunAggregationEvent.Message,
    STR2 := ',"lostEvents":');
CreateRunAggregationEvent.Message := CONCAT(STR1 := CreateRunAggregationEvent.Message,
    STR2 := UINT_TO_STRING(LostEventCount));
CreateRunAggregationEvent.Message := CONCAT(STR1 := CreateRunAggregationEvent.Message, STR2 := '}');

END_FUNCTION

// ---- Framework/EventBuffer/POU/EventBuffer.TcPOU
{region 'Documentation'}
(*!
<summary>Single-task event service. Initialize with static external event storage and status fields before use.</summary>
<description>
All producer and administrative calls use one PLC task; this service provides no concurrent-access synchronization. Bind one-based caller-owned storage of length 3..32767 and status fields before use; usable capacity is length minus one. Keep every binding alive and stable, and reinitialize after any online change. Publications never overwrite unread events. One logical consumer owns acknowledgements in each epoch. Sequence exhaustion is outside supported operation; the UDINT counter saturates rather than wrapping.
</description>
*)
{endregion}
FUNCTION_BLOCK INTERNAL EventBuffer IMPLEMENTS I_EventPublisher, I_EventBuffer
VAR
    EventFifo : Fifo;
    // Typed access for whole-array reset; valid only while the FIFO binding is valid.
    {attribute 'TcNoSymbol'}
    BufferEntries : POINTER TO ST_Event;
    EmptyEvent : ST_Event;
    BufferStatus : ST_EventBufferStatus;
    ReservedEntries : UINT;
    HasValidBinding : BOOL;
    {attribute 'TcNoSymbol'}
    FPublishedFifoControl : REFERENCE TO ST_FifoStatus;
    {attribute 'TcNoSymbol'}
    FPublishedStatus : REFERENCE TO ST_EventBufferStatus;
    FPublicationOnlineChangeCount : UDINT;
END_VAR

{region 'Documentation'}
(*!
<summary>Usable event positions, independent of occupancy and reservations; zero when invalid.</summary>
*)
{endregion}
{attribute 'monitoring' := 'call'}
PROPERTY PUBLIC Capacity : UINT //! Usable event positions, independent of occupancy and reservations; zero when invalid.
GET // PUBLIC
VAR
    CurrentFifoStatus : ST_FifoStatus;
END_VAR
Capacity := 0;
IF NOT IsValid THEN
    RETURN;
END_IF;
CurrentFifoStatus := FifoStatus;
Capacity := CurrentFifoStatus.BufferLength - 1;
END_GET
END_PROPERTY

{region 'Documentation'}
(*!
<summary>Release only eligible head events, bounded by the initial occupied entry count.</summary>
*)
{endregion}
METHOD PRIVATE DeleteBySequenceId
VAR_INPUT
    RequestedSequenceId : UDINT; //! Captured inclusive contiguous acknowledgement watermark for the current epoch; never a physical slot.
END_VAR
VAR
    CurrentFifoStatus : ST_FifoStatus;
    RemainingEntries : UINT;
    HeadEvent : ST_Event;
    ReadResult : INT;
    PopResult : INT;
END_VAR
CurrentFifoStatus := FifoStatus;
IF CurrentFifoStatus.ConfigError OR CurrentFifoStatus.IndexError THEN
    RETURN;
END_IF
IF RequestedSequenceId <= BufferStatus.DeletedSequenceId THEN
    RETURN;
END_IF
IF RequestedSequenceId > BufferStatus.SequenceId THEN
    PublishDeleteDiagnostic(Severity := E_EventSeverity.Warning,
        Reason := 'Requested sequence has not been produced.',
        RequestedSequenceId := RequestedSequenceId,
        HeadSequenceId := 0,
        FifoResult := TO_INT(E_FifoResult.NoTransfer));
    RETURN;
END_IF

FOR RemainingEntries := CurrentFifoStatus.ElementCount TO 1 BY -1 DO
    ReadResult := EventFifo.Read(Target := HeadEvent);
    IF ReadResult <= TO_INT(E_FifoResult.NoTransfer) THEN
        PublishDeleteDiagnostic(Severity := E_EventSeverity.Error,
            Reason := 'FIFO head could not be read.',
            RequestedSequenceId := RequestedSequenceId,
            HeadSequenceId := 0,
            FifoResult := ReadResult);
        RETURN;
    END_IF
    IF (HeadEvent.SequenceId = 0)
        OR (HeadEvent.SequenceId <= BufferStatus.DeletedSequenceId)
        OR (HeadEvent.SequenceId > RequestedSequenceId) THEN
        PublishDeleteDiagnostic(Severity := E_EventSeverity.Warning,
            Reason := 'FIFO head is outside the requested sequence range.',
            RequestedSequenceId := RequestedSequenceId,
            HeadSequenceId := HeadEvent.SequenceId,
            FifoResult := TO_INT(E_FifoResult.NoTransfer));
        RETURN;
    END_IF

    PopResult := EventFifo.Pop(Target := HeadEvent);
    IF PopResult <= TO_INT(E_FifoResult.NoTransfer) THEN
        IF PopResult <> TO_INT(E_FifoResult.NoTransfer) THEN
            PublishDeleteDiagnostic(Severity := E_EventSeverity.Error,
                Reason := 'FIFO could not remove and clear the head event.',
                RequestedSequenceId := RequestedSequenceId,
                HeadSequenceId := HeadEvent.SequenceId,
                FifoResult := PopResult);
        END_IF
        RETURN;
    END_IF

    BufferStatus.DeletedSequenceId := HeadEvent.SequenceId;
    IF BufferStatus.DeletedSequenceId >= RequestedSequenceId THEN
        EXIT;
    END_IF
END_FOR;

IF BufferStatus.DeletedSequenceId < RequestedSequenceId THEN
    PublishDeleteDiagnostic(Severity := E_EventSeverity.Warning,
        Reason := 'Buffer exhausted before the requested sequence was reached.',
        RequestedSequenceId := RequestedSequenceId,
        HeadSequenceId := 0,
        FifoResult := TO_INT(E_FifoResult.NoTransfer));
END_IF;
END_METHOD

{region 'Documentation'}
(*!
<summary>Value snapshot of readable-range metadata.</summary>
*)
{endregion}
{attribute 'monitoring' := 'variable'}
PROPERTY PUBLIC FifoStatus : ST_FifoStatus //! Value snapshot of readable-range metadata.
GET
FifoStatus := EventFifo.Status;
IF NOT HasValidBinding THEN
    FifoStatus.ConfigError := TRUE;
END_IF
END_GET
END_PROPERTY

{region 'Documentation'}
(*!
<summary>Usable free event positions before reservations; zero when invalid.</summary>
*)
{endregion}
{attribute 'monitoring' := 'call'}
PROPERTY PUBLIC FreeEntryCount : UINT //! Usable free event positions before reservations; zero when invalid.
GET
VAR
    CurrentFifoStatus : ST_FifoStatus;
END_VAR
FreeEntryCount := 0;
CurrentFifoStatus := FifoStatus;
IF CurrentFifoStatus.ConfigError OR CurrentFifoStatus.IndexError THEN
    RETURN;
END_IF
FreeEntryCount := CurrentFifoStatus.BufferLength - 1 - CurrentFifoStatus.ElementCount;
END_GET
END_PROPERTY

{region 'Documentation'}
(*!
<summary>Release only reservations, never events; FALSE changes neither count.</summary>
<description>
Requires an initialized valid binding, but no free capacity or valid FIFO indices.

Configuration and the owner contribution must be valid. Release is independent of free capacity and index validity; a zero release succeeds after the same accounting checks. It never removes events. Destructive buffer reset clears the aggregate count but does not repair stale owner-local contributions.
</description>
*)
{endregion}
METHOD PUBLIC FreeReservedSpace : BOOL //! TRUE after updating both reservation counts; FALSE leaves both unchanged.
VAR_INPUT
    EntryCount : UINT; //! Number of this owner's reserved entries to release; does not delete events.
END_VAR
VAR_IN_OUT
    OwnerReservedEntryCount : UINT; //! Owner's live reservation ledger; updated with the global count only on success, unchanged on rejection.
END_VAR
VAR
    CurrentFifoStatus : ST_FifoStatus;
END_VAR
FreeReservedSpace := FALSE;
CurrentFifoStatus := FifoStatus;
IF CurrentFifoStatus.ConfigError THEN
    RETURN;
END_IF
IF OwnerReservedEntryCount > ReservedEntries THEN
    RETURN;
END_IF
IF EntryCount > OwnerReservedEntryCount THEN
    RETURN;
END_IF

ReservedEntries := ReservedEntries - EntryCount;
OwnerReservedEntryCount := OwnerReservedEntryCount - EntryCount;
FreeReservedSpace := TRUE;
END_METHOD

{region 'Documentation'}
(*!
<summary>Read UTC Unix nanoseconds from the runtime's 100 ns system timestamp.</summary>
<description>
Source: Tc2_System.F_GetSystemTime, epoch 1601-01-01 UTC.

This is wall-clock publication time, not the ordering or acknowledgement identifier. Ordering and release use SequenceId independently of clock adjustments.
</description>
*)
{endregion}
METHOD PRIVATE GetUtcTimestamp : LINT //! UTC Unix time in nanoseconds converted from the 100 ns system timestamp.
VAR
    SystemTimeTicks : ULINT;
END_VAR
VAR CONSTANT
    UnixEpochOffsetTicks : LINT := 116444736000000000;
    NanosecondsPerTick : LINT := 100;
END_VAR
SystemTimeTicks := Tc2_System.F_GetSystemTime();
GetUtcTimestamp := (ULINT_TO_LINT(SystemTimeTicks) - UnixEpochOffsetTicks)
    * NanosecondsPerTick;
END_METHOD

{region 'Documentation'}
(*!
<summary>Bind one-based event storage and status fields; all storage must outlive this service.</summary>
<description>
FALSE publishes ConfigError and leaves the service unusable. Reinitialize after Online Change.

Buffer must have lower bound 1 and physical length 3..32767; usable capacity is one less. Success clears every entry and resets sequence, deletion, loss and aggregate reservations. A failed call invalidates the service and resets its internal counters; the old binding is not a recovery fallback. Call as part of full initialization with matching owner-ledger initialization, not as isolated recovery during execution.
</description>
*)
{endregion}
METHOD PUBLIC Initialize : BOOL //! TRUE when storage is bound and usable; FALSE leaves the service uninitialized.
VAR_IN_OUT
    Buffer : ARRAY[*] OF ST_Event; //! Caller-owned event array, bound by address until reinitialization; keep storage alive and unchanged.
    FifoControl : ST_FifoStatus; //! Caller-owned FIFO status storage, retained and updated after buffer operations; must outlive the service.
    Status : ST_EventBufferStatus; //! Caller-owned event-sequence/loss snapshot, retained and updated by the service; must outlive it.
END_VAR
Initialize := FALSE;
HasValidBinding := FALSE;
BufferEntries := 0;
FPublishedFifoControl REF= FifoControl;
FPublishedStatus REF= Status;
FPublicationOnlineChangeCount := TwinCAT_SystemInfoVarList._AppInfo.OnlineChangeCnt;
BufferStatus.SequenceId := 0;
BufferStatus.DeletedSequenceId := 0;
BufferStatus.LostEventCount := 0;
ReservedEntries := 0;

IF LOWER_BOUND(Buffer, 1) <> 1 THEN
    UpdatePublication();
    RETURN;
END_IF;
IF NOT EventFifo.Initialize(OverwriteIfFull := FALSE,
    Buffer := Buffer) THEN
    UpdatePublication();
    RETURN;
END_IF;

BufferEntries := ADR(Buffer[LOWER_BOUND(Buffer, 1)]);
HasValidBinding := TRUE;
Reset();
Initialize := IsValid;
END_METHOD

{region 'Documentation'}
(*!
<summary>FIFO binding, configuration and indices are valid.</summary>
*)
{endregion}
{attribute 'monitoring' := 'call'}
PROPERTY PUBLIC IsValid : BOOL //! FIFO binding, configuration and indices are valid.
GET
VAR
    CurrentFifoStatus : ST_FifoStatus;
END_VAR
CurrentFifoStatus := FifoStatus;
IsValid := NOT CurrentFifoStatus.ConfigError AND NOT CurrentFifoStatus.IndexError;
END_GET
END_PROPERTY

{region 'Documentation'}
(*!
<summary>Lost event count for producer diagnostics and aggregation.</summary>
*)
{endregion}
{attribute 'monitoring' := 'call'}
PROPERTY PUBLIC LostEventCount : UINT //! Lost event count for producer diagnostics and aggregation.
GET
LostEventCount := BufferStatus.LostEventCount;
END_GET
END_PROPERTY

{region 'Documentation'}
(*!
<summary>Process the captured release watermark; clear the caller&#x27;s field only if unchanged.</summary>
<description>
Zero is a no-op. Nonzero requests must belong to the current epoch and acknowledge all earlier unread events contiguously. Stale or future requests and inconsistent or unreachable heads are rejected or stop processing; partial deletion remains possible. The caller field is cleared when still equal to the snapshot even after rejection, so clearing alone does not prove deletion. Read Status.DeletedSequenceId for actual progress.
</description>
*)
{endregion}
METHOD PUBLIC ProcessDeleteRequest
VAR_IN_OUT
    SequenceId : UDINT; //! Inclusive deletion watermark; zero means no request. Cleared only if unchanged after processing.
END_VAR
VAR
    RequestedSequenceId : UDINT;
END_VAR
RequestedSequenceId := SequenceId;
IF RequestedSequenceId = 0 THEN
    RETURN;
END_IF

DeleteBySequenceId(RequestedSequenceId := RequestedSequenceId);
UpdatePublication();
IF SequenceId = RequestedSequenceId THEN
    SequenceId := 0;
END_IF
END_METHOD

{region 'Documentation'}
(*!
<summary>Store the capacity diagnostic without recursively generating another diagnostic.</summary>
*)
{endregion}
METHOD PRIVATE PublishCapacityWarning
VAR
    CapacityEvent : ST_Event;
END_VAR
CapacityEvent := EmptyEvent;
CapacityEvent.OwnerScope := E_OwnerScope.Framework;
CapacityEvent.EventType := E_EventType.Framework;
CapacityEvent.Severity := E_EventSeverity.Error;
CapacityEvent.Name := 'EventBuffer';
CapacityEvent.Message := 'UnitTest event buffer almost full. Further events may be lost.';
StoreEvent(Event := CapacityEvent);
END_METHOD

{region 'Documentation'}
(*!
<summary>Publish a bounded delete diagnostic with sequence context and the FIFO result.</summary>
*)
{endregion}
METHOD PRIVATE PublishDeleteDiagnostic
VAR_INPUT
    Severity : E_EventSeverity; //! Logging severity of the Framework diagnostic; independent of test Result.
    Reason : STRING(GVL_Constants.MessageLength); //! Reason text embedded with sequence context within the fixed diagnostic message capacity.
    RequestedSequenceId : UDINT; //! Captured acknowledgement watermark that could not be fully processed.
    HeadSequenceId : UDINT; //! Observed head event sequence, or zero when no head could be read.
    FifoResult : INT; //! FIFO transfer outcome included as diagnostic text; zero means no transfer.
END_VAR
VAR
    DiagnosticEvent : ST_Event;
END_VAR
DiagnosticEvent := EmptyEvent;
DiagnosticEvent.OwnerScope := E_OwnerScope.Framework;
DiagnosticEvent.EventType := E_EventType.Framework;
DiagnosticEvent.Severity := Severity;
DiagnosticEvent.Name := 'EventBuffer';
DiagnosticEvent.Message := CONCAT('Event-buffer delete: ', Reason);
DiagnosticEvent.Message := CONCAT(DiagnosticEvent.Message, ' Request=');
DiagnosticEvent.Message := CONCAT(DiagnosticEvent.Message, UDINT_TO_STRING(RequestedSequenceId));
DiagnosticEvent.Message := CONCAT(DiagnosticEvent.Message, ' Head=');
DiagnosticEvent.Message := CONCAT(DiagnosticEvent.Message, UDINT_TO_STRING(HeadSequenceId));
DiagnosticEvent.Message := CONCAT(DiagnosticEvent.Message, ' Deleted=');
DiagnosticEvent.Message := CONCAT(DiagnosticEvent.Message, UDINT_TO_STRING(BufferStatus.DeletedSequenceId));
DiagnosticEvent.Message := CONCAT(DiagnosticEvent.Message, ' Produced=');
DiagnosticEvent.Message := CONCAT(DiagnosticEvent.Message, UDINT_TO_STRING(BufferStatus.SequenceId));
DiagnosticEvent.Message := CONCAT(DiagnosticEvent.Message, ' FifoResult=');
DiagnosticEvent.Message := CONCAT(DiagnosticEvent.Message, INT_TO_STRING(FifoResult));
PublishEvent(Event := DiagnosticEvent);
END_METHOD

{region 'Documentation'}
(*!
<summary>Publish a value copy; positive slot on success, zero when full, negative on error.</summary>
<description>
Requires initialized storage. A capacity diagnostic never replaces the primary result.

The returned outcome belongs to the requested event. A successful insertion that leaves the ring almost full also attempts a Framework capacity diagnostic; that extra attempt may fail and increase LostEventCount without changing the primary return. Reservations do not block insertion or decrease on publication. Sequence numbers may therefore have gaps and loss makes the log incomplete.
</description>
*)
{endregion}
METHOD PUBLIC PublishEvent : INT //! Positive physical slot on success, zero when full, negative E_EventPublishResult on error.
VAR_INPUT
    Event : ST_Event; //! Event payload copied into the buffer; SequenceId and Timestamp are assigned by the publisher.
END_VAR
VAR
    CurrentFifoStatus : ST_FifoStatus;
END_VAR
PublishEvent := StoreEvent(Event := Event);
IF PublishEvent <= TO_INT(E_FifoResult.NoTransfer) THEN
    RETURN;
END_IF

CurrentFifoStatus := EventFifo.Status;
IF CurrentFifoStatus.BufferAlmostFull THEN
    PublishCapacityWarning();
END_IF
END_METHOD

{region 'Documentation'}
(*!
<summary>Aggregate producer reservations; not published externally.</summary>
*)
{endregion}
{attribute 'monitoring' := 'call'}
PROPERTY PUBLIC ReservedEntryCount : UINT //! Aggregate producer reservations; not published externally.
GET
ReservedEntryCount := ReservedEntries;
END_GET
END_PROPERTY

{region 'Documentation'}
(*!
<summary>Reserve additional event positions plus shared headroom; FALSE changes neither count.</summary>
<description>
Requires valid initialized configuration and a consistent owner contribution; positive requests also require valid indices.

For a positive EntryCount, physical free capacity must cover the updated aggregate reservation plus shared headroom. EntryCount zero succeeds after configuration and owner-contribution checks, without testing indices or headroom. Success updates both ledgers in one single-task call; no event or FIFO index changes. A failed call leaves both counts unchanged.
</description>
*)
{endregion}
METHOD PUBLIC ReserveSpace : BOOL //! TRUE after updating both reservation counts; FALSE leaves both unchanged.
VAR_INPUT
    EntryCount : UINT; //! Additional number of event entries to reserve for this owner.
    HeadroomEntryCount : UINT; //! Shared free entries checked for positive requests; not added to the owner's reservation.
END_VAR
VAR_IN_OUT
    OwnerReservedEntryCount : UINT; //! Owner's live reservation ledger; updated with the global count only on success, unchanged on rejection.
END_VAR
VAR
    CurrentFifoStatus : ST_FifoStatus;
    AvailableEntries : UINT;
    UpdatedReservedEntries : UDINT;
    RequiredFreeEntries : UDINT;
END_VAR
ReserveSpace := FALSE;
CurrentFifoStatus := FifoStatus;
IF CurrentFifoStatus.ConfigError THEN
    RETURN;
END_IF
IF OwnerReservedEntryCount > ReservedEntries THEN
    RETURN;
END_IF
IF EntryCount = 0 THEN
    ReserveSpace := TRUE;
    RETURN;
END_IF
IF CurrentFifoStatus.IndexError THEN
    RETURN;
END_IF

UpdatedReservedEntries := UINT_TO_UDINT(ReservedEntries) + UINT_TO_UDINT(EntryCount);
RequiredFreeEntries := UpdatedReservedEntries + UINT_TO_UDINT(HeadroomEntryCount);
AvailableEntries := CurrentFifoStatus.BufferLength - 1 - CurrentFifoStatus.ElementCount;
IF RequiredFreeEntries > UINT_TO_UDINT(AvailableEntries) THEN
    RETURN;
END_IF

ReservedEntries := UDINT_TO_UINT(UpdatedReservedEntries);
OwnerReservedEntryCount := UDINT_TO_UINT(UINT_TO_UDINT(OwnerReservedEntryCount)
    + UINT_TO_UDINT(EntryCount));
ReserveSpace := TRUE;
END_METHOD

{region 'Documentation'}
(*!
<summary>Clear bound storage and begin an empty epoch; binding must remain valid.</summary>
<description>
Does not access external commands and does not publish an event.

With a valid storage binding, clears the complete payload, FIFO state, sequence, deletion watermark, loss count and aggregate reservations. It does not rewrite owner-local ledgers. Run Control owns the preceding hierarchical release attempt and clearing external Reset/Delete commands. Consumers must discard acknowledgement assumptions from the old epoch. Invalid configuration prevents payload reset.
</description>
*)
{endregion}
METHOD PUBLIC Reset
VAR
    CurrentFifoStatus : ST_FifoStatus;
    EntryOffset : UINT;
END_VAR
CurrentFifoStatus := FifoStatus;
IF CurrentFifoStatus.ConfigError OR (BufferEntries = 0) THEN
    UpdatePublication();
    RETURN;
END_IF

FOR EntryOffset := 0 TO CurrentFifoStatus.BufferLength - 1 DO
    BufferEntries[EntryOffset] := EmptyEvent;
END_FOR
EventFifo.Reset();
BufferStatus.SequenceId := 0;
BufferStatus.DeletedSequenceId := 0;
BufferStatus.LostEventCount := 0;
ReservedEntries := 0;
UpdatePublication();
END_METHOD

{region 'Documentation'}
(*!
<summary>Value snapshot of sequence, deletion and loss status.</summary>
*)
{endregion}
{attribute 'monitoring' := 'variable'}
PROPERTY PUBLIC Status : ST_EventBufferStatus //! Value snapshot of sequence, deletion and loss status.
GET
Status := BufferStatus;
END_GET
END_PROPERTY

{region 'Documentation'}
(*!
<summary>Assign event identity/time and copy to FIFO; count each failed insertion once.</summary>
*)
{endregion}
METHOD PRIVATE StoreEvent : INT //! Positive physical slot on insertion, zero when full, negative E_EventPublishResult on error; failed insertion increments the saturating loss count.
VAR_IN_OUT
    Event : ST_Event; //! Borrowed payload whose SequenceId and Timestamp are assigned before the FIFO copy when a binding exists.
END_VAR
VAR CONSTANT
    MaximumSequenceId : UDINT := UDINT#16#FFFFFFFF;
    MaximumLostEventCount : UINT := UINT#16#FFFF;
END_VAR
IF NOT HasValidBinding THEN
    StoreEvent := TO_INT(E_FifoResult.ConfigError);
ELSE
    IF BufferStatus.SequenceId < MaximumSequenceId THEN
        BufferStatus.SequenceId := BufferStatus.SequenceId + 1;
    END_IF
    Event.SequenceId := BufferStatus.SequenceId;
    Event.Timestamp := GetUtcTimestamp();
    StoreEvent := EventFifo.Push(Data := Event);
END_IF

IF (StoreEvent <= TO_INT(E_FifoResult.NoTransfer))
    AND (BufferStatus.LostEventCount < MaximumLostEventCount) THEN
    BufferStatus.LostEventCount := BufferStatus.LostEventCount + 1;
END_IF

UpdatePublication();
END_METHOD

{region 'Documentation'}
(*!
<summary>Refresh only the bound producer-owned status fields; never copy the event array.</summary>
<description>
Do not dereference a publication binding from before an Online Change.
</description>
*)
{endregion}
METHOD PRIVATE UpdatePublication
IF NOT __ISVALIDREF(FPublishedFifoControl) OR NOT __ISVALIDREF(FPublishedStatus) THEN
    RETURN;
END_IF;
IF FPublicationOnlineChangeCount <> TwinCAT_SystemInfoVarList._AppInfo.OnlineChangeCnt THEN
    RETURN;
END_IF;

FPublishedFifoControl := FifoStatus;
FPublishedStatus := BufferStatus;
END_METHOD

END_FUNCTION_BLOCK

// ---- Framework/Common/Fifo/POU/Fifo.TcPOU
{region 'Documentation'}
(*!
<summary>Internal ST_Event ring buffer; storage stays owned by the caller.</summary>
<description>
Binds caller-owned ST_Event storage of physical length 3..32767; usable capacity is one less than that length. Logical transfer slots are one-based regardless of the array's declared lower bound. Keep the bound storage alive and unchanged. Any online change invalidates the binding and requires Initialize again. Reset discards logical contents without clearing payload bytes; Pop and Release clear transferred or acknowledged entries.


Transfer operations and positive-count Release check configuration before indices. Invalid indices cause those operations to reset both indices and return IndexError without transferring data; this discards logical contents without clearing old payloads. Status reports invalid state without repairing it. A zero-count Release is an unconditional no-op, including when uninitialized. Calls are serialized within one PLC task; this utility provides no synchronization.
</description>
*)
{endregion}
FUNCTION_BLOCK INTERNAL Fifo
VAR
    {attribute 'TcNoSymbol'}
    FBufferEntries : POINTER TO ST_Event;
    FBufferLength : UINT;
    FWriteIndex : UINT := 1;
    FReadIndex : UINT := 1;
    FInitialized : BOOL;
    FOverwriteOnFull : BOOL;
    {attribute 'TcNoSymbol'}
    FBindingOnlineChangeCount : UDINT;
END_VAR
VAR CONSTANT
    FirstBufferIndex : UINT := 1;
    MinimumBufferLength : UINT := 3;
    MaximumBufferLength : UINT := 32767;
    EmptyEvent : ST_Event := (SequenceId := 0);
END_VAR

{region 'Documentation'}
(*!
<summary>Check both logical indices before accessing bound storage.</summary>
*)
{endregion}
METHOD PRIVATE AreIndicesValid : BOOL //! TRUE when both stored logical indices are within 1..BufferLength.
AreIndicesValid := (FWriteIndex >= FirstBufferIndex) AND (FWriteIndex <= FBufferLength)
    AND (FReadIndex >= FirstBufferIndex) AND (FReadIndex <= FBufferLength);
END_METHOD

{region 'Documentation'}
(*!
<summary>Invalidate stored array access after instance relocation.</summary>
*)
{endregion}
METHOD FB_reinit : BOOL //! TRUE after invalidating the old array binding; Initialize is required before further access.
FInitialized := FALSE;
FBufferEntries := 0;
FBufferLength := 0;
FOverwriteOnFull := FALSE;
Reset();
FB_reinit := TRUE;
END_METHOD

{region 'Documentation'}
(*!
<summary>Bind live ST_Event storage; initialize indices without clearing the array.</summary>
<description>
The supplied array must contain 3..32767 entries and remain alive with a stable binding. One physical position stays unused. A failed call invalidates the previous binding. Initialize does not clear existing payload bytes.
</description>
*)
{endregion}
METHOD PUBLIC Initialize : BOOL //! TRUE when storage is bound and usable; FALSE leaves the service uninitialized.
VAR_INPUT
    OverwriteIfFull : BOOL := FALSE; //! TRUE replaces the oldest event when full; default FALSE rejects insertion.
END_VAR
VAR_IN_OUT
    Buffer : ARRAY[*] OF ST_Event; //! Caller-owned event array, bound by address until reinitialization; keep storage alive and unchanged.
END_VAR
VAR
    ConfiguredBufferLength : LINT;
END_VAR
Initialize := FALSE;
FInitialized := FALSE;
FBufferEntries := 0;
FBufferLength := 0;
FOverwriteOnFull := FALSE;
Reset();

ConfiguredBufferLength := TO_LINT(UPPER_BOUND(Buffer, 1))
    - TO_LINT(LOWER_BOUND(Buffer, 1)) + 1;
IF (ConfiguredBufferLength < TO_LINT(MinimumBufferLength))
    OR (ConfiguredBufferLength > TO_LINT(MaximumBufferLength)) THEN
    RETURN;
END_IF;

FBufferEntries := ADR(Buffer[LOWER_BOUND(Buffer, 1)]);
FBufferLength := LINT_TO_UINT(ConfiguredBufferLength);
FOverwriteOnFull := OverwriteIfFull;
FBindingOnlineChangeCount := TwinCAT_SystemInfoVarList._AppInfo.OnlineChangeCnt;
FInitialized := TRUE;
Initialize := TRUE;
END_METHOD

{region 'Documentation'}
(*!
<summary>Validate binding lifetime and capacity without dereferencing the array.</summary>
*)
{endregion}
METHOD PRIVATE IsConfigValid : BOOL //! TRUE when initialization, capacity and binding are valid and no online change has invalidated the binding.
IsConfigValid := FInitialized AND (FBufferEntries <> 0)
    AND (FBufferLength >= MinimumBufferLength) AND (FBufferLength <= MaximumBufferLength)
    AND (FBindingOnlineChangeCount = TwinCAT_SystemInfoVarList._AppInfo.OnlineChangeCnt);
END_METHOD

{region 'Documentation'}
(*!
<summary>Reject output storage overlapping the array; requires valid configuration.</summary>
*)
{endregion}
METHOD PRIVATE IsOutputTargetValid : BOOL //! TRUE when Target does not overlap bound event storage; configuration must already be valid.
VAR_IN_OUT CONSTANT
    Target : ST_Event; //! Borrowed output object whose address range is checked against the bound event array.
END_VAR
VAR
    TargetStart : __UXINT;
    BufferStart : __UXINT;
    BufferEnd : __UXINT;
END_VAR
TargetStart := TO___UXINT(ADR(Target));
BufferStart := TO___UXINT(FBufferEntries);
BufferEnd := TO___UXINT(ADR(FBufferEntries[FBufferLength - 1]))
    + TO___UXINT(SIZEOF(ST_Event) - 1);
IF TargetStart < BufferStart THEN
    IsOutputTargetValid := (BufferStart - TargetStart) >= TO___UXINT(SIZEOF(ST_Event));
ELSE
    IsOutputTargetValid := TargetStart > BufferEnd;
END_IF;
END_METHOD

{region 'Documentation'}
(*!
<summary>Advance one logical slot, wrapping before incrementing past capacity.</summary>
*)
{endregion}
METHOD PRIVATE NextIndex : UINT //! Following one-based ring index, wrapping from BufferLength to 1.
VAR_INPUT
    CurrentIndex : UINT; //! Caller-validated logical ring index in 1..BufferLength.
END_VAR
IF CurrentIndex = FBufferLength THEN
    NextIndex := FirstBufferIndex;
ELSE
    NextIndex := CurrentIndex + 1;
END_IF;
END_METHOD

{region 'Documentation'}
(*!
<summary>Copy and remove the oldest event; Target must be outside the bound array.</summary>
*)
{endregion}
METHOD PUBLIC Pop : INT //! Positive physical slot on transfer, zero when no transfer is possible, negative E_FifoResult on error.
VAR_IN_OUT
    Target : ST_Event; //! Destination for the oldest event copy; must not overlap the bound array.
END_VAR
IF NOT IsConfigValid() THEN
    Pop := TO_INT(E_FifoResult.ConfigError);
    RETURN;
END_IF;
IF NOT AreIndicesValid() THEN
    Reset();
    Pop := TO_INT(E_FifoResult.IndexError);
    RETURN;
END_IF;
IF FReadIndex = FWriteIndex THEN
    Pop := TO_INT(E_FifoResult.NoTransfer);
    RETURN;
END_IF;
IF NOT IsOutputTargetValid(Target := Target) THEN
    Pop := TO_INT(E_FifoResult.DataError);
    RETURN;
END_IF;

Target := FBufferEntries[FReadIndex - FirstBufferIndex];
FBufferEntries[FReadIndex - FirstBufferIndex] := EmptyEvent;
Pop := UINT_TO_INT(FReadIndex);
FReadIndex := NextIndex(CurrentIndex := FReadIndex);
END_METHOD

{region 'Documentation'}
(*!
<summary>Copy one event; return its physical slot, no transfer, or a named error.</summary>
*)
{endregion}
METHOD PUBLIC Push : INT //! Positive physical slot on transfer, zero when no transfer is possible, negative E_FifoResult on error.
VAR_INPUT
    Data : ST_Event; //! Event copied into the next free FIFO slot.
END_VAR
VAR
    NextWriteIndex : UINT;
    BufferFull : BOOL;
END_VAR
IF NOT IsConfigValid() THEN
    Push := TO_INT(E_FifoResult.ConfigError);
    RETURN;
END_IF;
IF NOT AreIndicesValid() THEN
    Reset();
    Push := TO_INT(E_FifoResult.IndexError);
    RETURN;
END_IF;

NextWriteIndex := NextIndex(CurrentIndex := FWriteIndex);
BufferFull := NextWriteIndex = FReadIndex;
IF BufferFull AND NOT FOverwriteOnFull THEN
    Push := TO_INT(E_FifoResult.NoTransfer);
    RETURN;
END_IF;

FBufferEntries[FWriteIndex - FirstBufferIndex] := Data;
Push := UINT_TO_INT(FWriteIndex);
IF BufferFull THEN
    FReadIndex := NextIndex(CurrentIndex := FReadIndex);
END_IF;
FWriteIndex := NextWriteIndex;
END_METHOD

{region 'Documentation'}
(*!
<summary>Copy without removing the oldest event; Target must be outside the bound array.</summary>
*)
{endregion}
METHOD PUBLIC Read : INT //! Positive physical slot on transfer, zero when no transfer is possible, negative E_FifoResult on error.
VAR_IN_OUT
    Target : ST_Event; //! Destination for the oldest event copy; must not overlap the bound array.
END_VAR
IF NOT IsConfigValid() THEN
    Read := TO_INT(E_FifoResult.ConfigError);
    RETURN;
END_IF;
IF NOT AreIndicesValid() THEN
    Reset();
    Read := TO_INT(E_FifoResult.IndexError);
    RETURN;
END_IF;
IF FReadIndex = FWriteIndex THEN
    Read := TO_INT(E_FifoResult.NoTransfer);
    RETURN;
END_IF;
IF NOT IsOutputTargetValid(Target := Target) THEN
    Read := TO_INT(E_FifoResult.DataError);
    RETURN;
END_IF;

Target := FBufferEntries[FReadIndex - FirstBufferIndex];
Read := UINT_TO_INT(FReadIndex);
END_METHOD

{region 'Documentation'}
(*!
<summary>Clear and release Count oldest entries; an excessive count changes nothing.</summary>
<description>
Count zero returns NoTransfer before configuration or index checks. For a positive count, configuration/index validation precedes the occupancy-range check. A valid excessive request returns ReleaseCountError without mutation; an index error instead resets logical contents and returns IndexError. Clearing a valid range costs proportionally to Count.
</description>
*)
{endregion}
METHOD PUBLIC Release : INT //! Number of released entries; negative E_FifoResult on failure.
VAR_INPUT
    Count : UINT; //! Number of oldest events to clear and release; excessive requests change nothing.
END_VAR
VAR
    AvailableCount : UINT;
    ReleaseReadIndex : UINT;
    ClearedCount : UINT;
END_VAR
IF Count = 0 THEN
    Release := TO_INT(E_FifoResult.NoTransfer);
    RETURN;
END_IF;
IF NOT IsConfigValid() THEN
    Release := TO_INT(E_FifoResult.ConfigError);
    RETURN;
END_IF;
IF NOT AreIndicesValid() THEN
    Reset();
    Release := TO_INT(E_FifoResult.IndexError);
    RETURN;
END_IF;

IF FWriteIndex >= FReadIndex THEN
    AvailableCount := FWriteIndex - FReadIndex;
ELSE
    AvailableCount := FBufferLength - FReadIndex + FWriteIndex;
END_IF;
IF Count > AvailableCount THEN
    Release := TO_INT(E_FifoResult.ReleaseCountError);
    RETURN;
END_IF;

ReleaseReadIndex := FReadIndex;
FOR ClearedCount := FirstBufferIndex TO Count DO
    FBufferEntries[ReleaseReadIndex - FirstBufferIndex] := EmptyEvent;
    ReleaseReadIndex := NextIndex(CurrentIndex := ReleaseReadIndex);
END_FOR;

FReadIndex := ReleaseReadIndex;
Release := UINT_TO_INT(Count);
END_METHOD

{region 'Documentation'}
(*!
<summary>Discard logical contents, retaining binding and payload storage.</summary>
*)
{endregion}
METHOD PUBLIC Reset
FWriteIndex := FirstBufferIndex;
FReadIndex := FirstBufferIndex;
END_METHOD

{region 'Documentation'}
(*!
<summary>Snapshot of binding validity, indices and derived occupancy.</summary>
*)
{endregion}
PROPERTY PUBLIC Status : ST_FifoStatus //! Snapshot of binding validity, indices and derived occupancy.
GET
Status.ConfigError := NOT IsConfigValid();
Status.IndexError := FALSE;
Status.IndexIn := FWriteIndex;
Status.IndexOut := FReadIndex;
Status.BufferAlmostFull := FALSE;
Status.BufferFull := FALSE;
Status.BufferEmpty := FALSE;
Status.ElementCount := 0;
Status.BufferLength := FBufferLength;
IF Status.ConfigError THEN
    RETURN;
END_IF

Status.IndexError := NOT AreIndicesValid();
IF Status.IndexError THEN
    RETURN;
END_IF

IF FWriteIndex >= FReadIndex THEN
    Status.ElementCount := FWriteIndex - FReadIndex;
ELSE
    Status.ElementCount := FBufferLength - FReadIndex + FWriteIndex;
END_IF
Status.BufferEmpty := Status.ElementCount = 0;
Status.BufferAlmostFull := Status.ElementCount = FBufferLength - 2;
Status.BufferFull := Status.ElementCount >= FBufferLength - 1;
END_GET
END_PROPERTY

END_FUNCTION_BLOCK

// ---- Framework/Common/POU/IsNameValid.TcPOU
{region 'Documentation'}
(*!
<summary>Validates the unshortened full name against hierarchy, character and length rules. Depth: 1 Run Control, 2 Suite, 3 Test Case, 4 Assertion (remaining suffix may contain dots).</summary>
*)
{endregion}
FUNCTION INTERNAL IsNameValid : BOOL //! TRUE only when the full name satisfies depth, ASCII character and length rules.
VAR_INPUT
    Depth : UINT; //! Required hierarchy depth: 1 Run Control, 2 Suite, 3 Test Case, 4 Assertion.
END_VAR
VAR_IN_OUT CONSTANT
    Name : STRING(2 * GVL_Constants.NameLength + 1); //! Unshortened full hierarchical name; borrowed read-only and checked against Depth and NameLength.
END_VAR
VAR
    Index : INT;
    NameLength : INT;
    Segment : UINT := 1;
    SegmentLength : UINT;
    Character : BYTE;
END_VAR
VAR CONSTANT
    RootDepth : UINT := 1;
    AssertionDepth : UINT := 4;
    HierarchySeparator : BYTE := 16#2E;
    FirstUppercaseLetter : BYTE := 16#41;
    LastUppercaseLetter : BYTE := 16#5A;
    FirstLowercaseLetter : BYTE := 16#61;
    LastLowercaseLetter : BYTE := 16#7A;
    FirstDigit : BYTE := 16#30;
    LastDigit : BYTE := 16#39;
    Underscore : BYTE := 16#5F;
    Hyphen : BYTE := 16#2D;
    LastAsciiCharacter : BYTE := 16#7F;
END_VAR

IsNameValid := FALSE;
NameLength := LEN(Name);
IF (NameLength = 0) OR (NameLength > GVL_Constants.NameLength) THEN
    RETURN;
END_IF;

IF (Depth < RootDepth) OR (Depth > AssertionDepth) THEN
    RETURN;
END_IF;

FOR Index := 0 TO NameLength - 1 DO
    // SA0175: ASCII name contract; byte-based access is intentional and bounded.
    {analysis -175}
    Character := Name[Index];
    {analysis +175}
    IF (Depth = AssertionDepth) AND (Segment = AssertionDepth) THEN
        IF Character > LastAsciiCharacter THEN
            RETURN;
        END_IF;
        SegmentLength := SegmentLength + 1;
    ELSIF Character = HierarchySeparator THEN
        IF (SegmentLength = 0) OR (Segment >= Depth) THEN
            RETURN;
        END_IF;
        Segment := Segment + 1;
        SegmentLength := 0;
    ELSE
        IF NOT (((Character >= FirstUppercaseLetter) AND (Character <= LastUppercaseLetter))
            OR ((Character >= FirstLowercaseLetter) AND (Character <= LastLowercaseLetter))
            OR ((Character >= FirstDigit) AND (Character <= LastDigit))
            OR (Character = Underscore) OR (Character = Hyphen)) THEN
            RETURN;
        END_IF;
        SegmentLength := SegmentLength + 1;
    END_IF;
END_FOR;

IsNameValid := (Segment = Depth) AND (SegmentLength > 0);

END_FUNCTION

// ---- Framework/EventBuffer/POU/TriggerEvents/CreateResetEvent.TcPOU
{region 'Documentation'}
(*!
<summary>Constructs a reset trigger event without publishing it.</summary>
<description>
The caller supplies valid ASCII owner context; publication assigns sequence and time.
</description>
*)
{endregion}
FUNCTION CreateResetEvent : ST_Event //! Constructed event value; not published. The publisher assigns SequenceId and Timestamp.
VAR_INPUT
    OwnerScope : E_OwnerScope; //! Semantic owner category recorded in the event.
    Name : STRING(GVL_Constants.NameLength); //! Hierarchical owner name used to identify events; must satisfy the naming contract.
    ResourceName : STRING(GVL_Constants.ResourceNameLength) := ''; //! Optional resource context for diagnostics; empty by default.
    State : E_State; //! Owner lifecycle state recorded in the event.
END_VAR

CreateResetEvent.SequenceId := 0;
CreateResetEvent.Timestamp := 0;
CreateResetEvent.OwnerScope := OwnerScope;
CreateResetEvent.EventType := E_EventType.Trigger;
CreateResetEvent.Severity := E_EventSeverity.Info;
CreateResetEvent.Name := Name;
CreateResetEvent.ResourceName := ResourceName;
CreateResetEvent.State := State;
CreateResetEvent.Result := E_Result.NotEvaluated;
CreateResetEvent.Message := 'Reset trigger.';

END_FUNCTION

// ---- Framework/EventBuffer/POU/TriggerEvents/CreateAbortEvent.TcPOU
{region 'Documentation'}
(*!
<summary>Constructs an abort trigger event without publishing it.</summary>
<description>
The caller supplies valid ASCII owner context; publication assigns sequence and time.
</description>
*)
{endregion}
FUNCTION CreateAbortEvent : ST_Event //! Constructed event value; not published. The publisher assigns SequenceId and Timestamp.
VAR_INPUT
    OwnerScope : E_OwnerScope; //! Semantic owner category recorded in the event.
    Name : STRING(GVL_Constants.NameLength); //! Hierarchical owner name used to identify events; must satisfy the naming contract.
    ResourceName : STRING(GVL_Constants.ResourceNameLength) := ''; //! Optional resource context for diagnostics; empty by default.
    State : E_State; //! Owner lifecycle state recorded in the event.
END_VAR

CreateAbortEvent.SequenceId := 0;
CreateAbortEvent.Timestamp := 0;
CreateAbortEvent.OwnerScope := OwnerScope;
CreateAbortEvent.EventType := E_EventType.Trigger;
CreateAbortEvent.Severity := E_EventSeverity.Info;
CreateAbortEvent.Name := Name;
CreateAbortEvent.ResourceName := ResourceName;
CreateAbortEvent.State := State;
CreateAbortEvent.Result := E_Result.NotEvaluated;
CreateAbortEvent.Message := 'Abort trigger.';

END_FUNCTION

// ---- Framework/EventBuffer/POU/TriggerEvents/CreateStartEvent.TcPOU
{region 'Documentation'}
(*!
<summary>Constructs a start trigger event without publishing it.</summary>
<description>
The caller supplies valid ASCII owner context; publication assigns sequence and time.
</description>
*)
{endregion}
FUNCTION CreateStartEvent : ST_Event //! Constructed event value; not published. The publisher assigns SequenceId and Timestamp.
VAR_INPUT
    OwnerScope : E_OwnerScope; //! Semantic owner category recorded in the event.
    Name : STRING(GVL_Constants.NameLength); //! Hierarchical owner name used to identify events; must satisfy the naming contract.
    ResourceName : STRING(GVL_Constants.ResourceNameLength) := ''; //! Optional resource context for diagnostics; empty by default.
    State : E_State; //! Owner lifecycle state recorded in the event.
END_VAR

CreateStartEvent.SequenceId := 0;
CreateStartEvent.Timestamp := 0;
CreateStartEvent.OwnerScope := OwnerScope;
CreateStartEvent.EventType := E_EventType.Trigger;
CreateStartEvent.Severity := E_EventSeverity.Info;
CreateStartEvent.Name := Name;
CreateStartEvent.ResourceName := ResourceName;
CreateStartEvent.State := State;
CreateStartEvent.Result := E_Result.NotEvaluated;
CreateStartEvent.Message := 'Start trigger.';

END_FUNCTION

// ---- SelfTests/TestSuites/TestSuite_Smoke.TcPOU
{region 'Documentation'}
(*!
<summary>Runs the single successful smoke Test Case through the production Suite lifecycle.</summary>
*)
{endregion}
FUNCTION_BLOCK TestSuite_Smoke EXTENDS TestSuiteBase
VAR
    FSmoke : Test_Smoke;
    FTestCases : ARRAY[1..TestCaseCapacity] OF I_TestCase;
END_VAR
VAR CONSTANT
    TestCaseCapacity : UINT := 1;
END_VAR

SUPER^();

{region 'Documentation'}
(*!
<summary>Initializes the smoke Test Case and registers it for serial execution.</summary>
*)
{endregion}
METHOD PROTECTED Configure
VAR_IN_OUT
    // SA0167: Borrowed builder; VAR_IN_OUT creates no temporary instance.
    {attribute 'analysis' := '-167'}
    Builder : TestSuiteConfigurationBuilder; //! Borrowed owner configuration builder used only during this Configure call; register this owner's concrete children.
END_VAR
VAR
    TestConfig : ST_TestCaseConfig;
END_VAR
Builder.Initialize(Mode := E_OrchestrationMode.Serial,
    TestCases := FTestCases);

FSmoke.Initialize(Parent := THIS^,
    TestName := 'Execution',
    Config := TestConfig);
Builder.Register(TestCase := FSmoke);
END_METHOD

{region 'Documentation'}
(*!
<summary>Returns the registered Test Case from the same array used during configuration.</summary>
*)
{endregion}
METHOD PUBLIC GetTestCase : I_TestCase //! Typed child interface at the original array index; zero when no entry is available.
VAR_INPUT
    Index : DINT; //! Original occupied child-array index, rather than an ordinal position.
END_VAR
GetTestCase := 0;
IF (ChildCount = 0) OR (Index < ChildArrayLowerBound)
    OR (DINT_TO_LINT(Index) >= DINT_TO_LINT(ChildArrayLowerBound) + UINT_TO_LINT(ChildCount)) THEN
    RETURN;
END_IF;

GetTestCase := FTestCases[Index];
END_METHOD

{region 'Documentation'}
(*!
<summary>Calls the owned Test Case once per initialized Suite cycle, including completion.</summary>
*)
{endregion}
METHOD PROTECTED ProcessTestCases
FSmoke();
END_METHOD

END_FUNCTION_BLOCK

// ---- Framework/TestSuites/POU/TestSuiteBase.TcPOU
{region 'Documentation'}
(*!
<summary>Base-owned Suite lifecycle and orchestration of a concrete Test Case collection.</summary>
<description>
The Run Control calls Initialize. Implement Configure, GetTestCase and ProcessTestCases; the
concrete FB body calls SUPER^() once per task cycle.

Configure initializes and registers static children. The base owns builder finalization,
Orchestrator initialization and execution, timeouts, aggregation and owner events. Continue calling
every child during Completing and Completed; finalized owner results remain held while status is
refreshed.
</description>
*)
{endregion}
FUNCTION_BLOCK ABSTRACT TestSuiteBase IMPLEMENTS I_TestSuite, I_OrchestratableCollection
VAR
    /// Instance binding; derived test adapters may assign it before first use.
    FEventPublisher : I_EventPublisher;
    FName : STRING(GVL_Constants.NameLength);
    FResourceName : STRING(GVL_Constants.ResourceNameLength);
    FConfig : ST_TestSuiteConfig;
    FCollectionConfiguration : ST_TestCaseCollectionConfig;
    FInitialized : BOOL;
    FHasTimeout : BOOL;
    FHasResetTimeout : BOOL;
    FHasAbortTimeout : BOOL;
    FCheckingInitialization : BOOL;
    FConfigError : BOOL;
    FOrchestrator : I_Orchestrator;
    FDefaultOrchestrator : Orchestrator;
    FStatus : ST_TestSuiteStatus;
    FResult : E_Result := E_Result.NotEvaluated;
    FMethodRequests : ST_Command;
    FState : E_State := E_State.Uninitialized;
    FExecutionTimer : Stopwatch;
    FStateTimer : Stopwatch;
    FAggregator : ResultAggregator;
    FTestCaseCountInactive : UINT;
    FTestCaseCountIdle : UINT;
    FTestCaseCountRunning : UINT;
    FTestCaseCountCompleted : UINT;
    FTestCaseCountError : UINT;
    FCollectionValid : BOOL;
    FChildrenError : BOOL;
    FChildrenAborted : BOOL;
    FChildrenCompleted : BOOL;
    FChildrenAbortFinished : BOOL;
    FExecutionSlot : UINT;
    FReservedEntryCount : UINT;
END_VAR
VAR_TEMP
    Requests : ST_Command;
    OrchestratorTask : E_OrchestratorTask;
END_VAR

ProcessRequests(InputRequests := FMethodRequests, Requests => Requests);

FExecutionTimer.Update();
FStateTimer.Update();

Sequencer(Requests := Requests);

IF IsInitialized THEN
    OrchestratorTask := MapOrchestratorTask(State := FState,
        CurrentTask := FOrchestrator.CurrentTask);
    FOrchestrator.Execute(Task := OrchestratorTask);

    ProcessTestCases();
    AggregateResults();
END_IF;

UpdateResult();
UpdateStatus();
EmitFinalizationEvents();

{region 'Documentation'}
(*!
<summary>Aggregates results and execution counters after child calls; refreshes observations from the same snapshots.</summary>
*)
{endregion}
METHOD PRIVATE AggregateResults
VAR
    Count : UINT;
    FirstIndex : DINT;
    LastIndex : DINT;
    Index : LINT;
    ChildStatus : ST_TestCaseStatus;
    ChildResult : E_Result;
END_VAR
Count := ChildCount;
FTestCaseCountInactive := 0;
FTestCaseCountIdle := 0;
FTestCaseCountRunning := 0;
FTestCaseCountCompleted := 0;
FTestCaseCountError := 0;
FAggregator.Reset();
FCollectionValid := FALSE;
FChildrenCompleted := FALSE;
FChildrenAbortFinished := FALSE;
FChildrenError := FALSE;
FChildrenAborted := FALSE;

IF NOT FInitialized OR (Count = 0) THEN
    RETURN;
END_IF;
FirstIndex := ChildArrayLowerBound;
LastIndex := ChildArrayUpperBound;
IF DINT_TO_LINT(LastIndex) - DINT_TO_LINT(FirstIndex) + 1 < UINT_TO_LINT(Count) THEN
    RETURN;
END_IF;

FCollectionValid := TRUE;
FChildrenCompleted := TRUE;
FChildrenAbortFinished := TRUE;
FOR Index := DINT_TO_LINT(FirstIndex) TO DINT_TO_LINT(FirstIndex) + UINT_TO_LINT(Count) - 1 DO
    IF NOT ObserveTestCase(Child := GetTestCase(Index := LINT_TO_DINT(Index)),
        ChildStatus => ChildStatus) THEN
        FTestCaseCountError := FTestCaseCountError + 1;
        FAggregator.AddResult(Result := E_Result.Error);
        CONTINUE;
    END_IF;

    ChildResult := ChildStatus.Execution.Result;
    CASE ChildResult OF
        E_Result.NotEvaluated, E_Result.Passed, E_Result.Failed, E_Result.Abort, E_Result.Error:
            FAggregator.AddResult(Result := ChildResult);
    ELSE
        ChildResult := E_Result.Error;
        FAggregator.AddResult(Result := ChildResult);
    END_CASE;

    CASE ChildStatus.Execution.ExecutionStatus OF
        E_ExecutionStatus.Inactive:
            FTestCaseCountInactive := FTestCaseCountInactive + 1;
        E_ExecutionStatus.Idle:
            FTestCaseCountIdle := FTestCaseCountIdle + 1;
        E_ExecutionStatus.Running:
            FTestCaseCountRunning := FTestCaseCountRunning + 1;
        E_ExecutionStatus.Completed:
            FTestCaseCountCompleted := FTestCaseCountCompleted + 1;
    ELSE
        // Transitional execution states have no dedicated counter in the status contract.
    END_CASE;
    IF (ChildStatus.Execution.ExecutionStatus = E_ExecutionStatus.Error) OR (ChildResult = E_Result.Error) THEN
        FTestCaseCountError := FTestCaseCountError + 1;
    END_IF;

END_FOR;
END_METHOD

{region 'Documentation'}
(*!
<summary>Applies permitted transitions; rejection holds state/timers and emits phase-dependent diagnostics or latches Error.</summary>
*)
{endregion}
METHOD PRIVATE ChangeState
VAR_INPUT
    NewState : E_State; //! Requested lifecycle destination; identical state is a no-op and rejection leaves state and timers unchanged.
END_VAR
IF NewState = FState THEN
    RETURN;
END_IF;
IF NOT IsStateTransitionAllowed(NewState := NewState) THEN
    CASE FState OF
        E_State.Uninitialized:
            RETURN;

        E_State.Completed:
            PublishEvent(Event := CreateInvalidStateTransitionEvent(OwnerScope := E_OwnerScope.TestSuite,
                Name := FName,
                ResourceName := FResourceName,
                StateOld := FState,
                StateNew := NewState));
    ELSE
        IF FResult <> E_Result.Error THEN
            PublishEvent(Event := CreateInvalidStateTransitionEvent(OwnerScope := E_OwnerScope.TestSuite,
                Name := FName,
                ResourceName := FResourceName,
                StateOld := FState,
                StateNew := NewState));
        END_IF;
        FResult := E_Result.Error;
    END_CASE;
    RETURN;
END_IF;

CASE NewState OF
    E_State.Uninitialized:
        FExecutionTimer.Reset();
        FStateTimer.Start();
        FResult := E_Result.NotEvaluated;
    E_State.Reset:
        FHasTimeout := FALSE;
        FHasResetTimeout := FALSE;
        FHasAbortTimeout := FALSE;
        IF (FState = E_State.Starting) OR (FState = E_State.Running) OR (FState = E_State.Completing)
            OR (FState = E_State.Aborting) OR (FState = E_State.AbortingFromError) THEN
            PublishEvent(Event := CreateResetWarningEvent(OwnerScope := E_OwnerScope.TestSuite,
                Name := FName,
                ResourceName := FResourceName,
                State := FState));
        END_IF;
        FExecutionTimer.Reset();
        FStateTimer.Start();
        FResult := E_Result.NotEvaluated;
    E_State.Idle:
        FStateTimer.Start();
    E_State.Starting:
        FStateTimer.Start();
        FExecutionTimer.Start();
    E_State.Running:
        FStateTimer.Start();
    E_State.Completing:
        FExecutionTimer.Stop();
        FStateTimer.Start();
    E_State.Completed:
        FStateTimer.Start();
    E_State.Aborting:
        FExecutionTimer.Stop();
        FStateTimer.Start();
        IF FResult <> E_Result.Error THEN
            FResult := E_Result.Abort;
        END_IF;
    E_State.AbortingFromError:
        FExecutionTimer.Stop();
        IF FState <> E_State.Aborting THEN
            FStateTimer.Start();
        END_IF;
        FResult := E_Result.Error;
ELSE
    RETURN;
END_CASE;
PublishEvent(Event := CreateStateTransitionEvent(OwnerScope := E_OwnerScope.TestSuite,
    Name := FName,
    ResourceName := FResourceName,
    StateOld := FState,
    StateNew := NewState));
FState := NewState;
END_METHOD

{region 'Documentation'}
(*!
<summary>Validates timeouts, the initialized Orchestrator and every registered child.</summary>
<description>
Called after builder finalization and helper initialization. An override must include
SUPER^.CheckInitialization(), preserve failure and check any additional application setup.

Timeout, ResetTimeout and AbortTimeout must be positive. The base reports its first failed
check; FALSE prevents successful initialization.
</description>
*)
{endregion}
METHOD PROTECTED CheckInitialization : BOOL //! TRUE when the configured setup is valid; FALSE reports invalid setup and prevents initialization.
VAR
    Index : LINT;
    Child : I_TestCase;
END_VAR
CheckInitialization := FALSE;
IF (FConfig.Timeout = T#0ms) OR (FConfig.ResetTimeout = T#0ms) OR (FConfig.AbortTimeout = T#0ms) THEN
    PublishInitializationError(Message := 'Suite timeouts must be greater than zero.');
    RETURN;
END_IF;
IF NOT FOrchestrator.IsInitialized THEN
    PublishInitializationError(Message := 'Orchestrator initialization is invalid.');
    RETURN;
END_IF;
IF (ChildCount = 0)
    OR (DINT_TO_LINT(ChildArrayUpperBound) - DINT_TO_LINT(ChildArrayLowerBound) + 1 < UINT_TO_LINT(ChildCount)) THEN
    PublishInitializationError(Message := 'Invalid registered Test Case range.');
    RETURN;
END_IF;
FOR Index := DINT_TO_LINT(ChildArrayLowerBound) TO DINT_TO_LINT(ChildArrayLowerBound) + UINT_TO_LINT(ChildCount) - 1 DO
    Child := GetTestCase(Index := LINT_TO_DINT(Index));
    IF Child = 0 THEN
        PublishInitializationError(Message := CONCAT('Missing Test Case at index ', LINT_TO_STRING(Index)));
        RETURN;
    END_IF;
    IF NOT Child.IsInitialized THEN
        PublishInitializationError(Message := CONCAT('Test Case is not initialized: ', Child.Name));
        RETURN;
    END_IF;
END_FOR;
CheckInitialization := TRUE;
END_METHOD

{region 'Documentation'}
(*!
<summary>Actual array lower bound; zero when no configuration is available.</summary>
*)
{endregion}
{attribute 'monitoring' := 'call'}
PROPERTY PUBLIC ChildArrayLowerBound : DINT //! Actual array lower bound; zero when no configuration is available.
GET // PUBLIC
ChildArrayLowerBound := 0;
IF NOT (FInitialized OR FCheckingInitialization) OR NOT FCollectionConfiguration.IsValid THEN
    RETURN;
END_IF;
ChildArrayLowerBound := FCollectionConfiguration.FirstIndex;
END_GET
END_PROPERTY

{region 'Documentation'}
(*!
<summary>Actual array upper bound, including unused capacity; process only ChildCount
entries.</summary>
*)
{endregion}
{attribute 'monitoring' := 'call'}
PROPERTY PUBLIC ChildArrayUpperBound : DINT //! Actual array upper bound, including unused capacity; process only ChildCount entries.
GET // PUBLIC
ChildArrayUpperBound := 0;
IF NOT (FInitialized OR FCheckingInitialization) OR NOT FCollectionConfiguration.IsValid THEN
    RETURN;
END_IF;
ChildArrayUpperBound := FCollectionConfiguration.LastIndex;
END_GET
END_PROPERTY

{region 'Documentation'}
(*!
<summary>Registered population starting at ChildArrayLowerBound; zero when unavailable.</summary>
*)
{endregion}
{attribute 'monitoring' := 'call'}
PROPERTY PUBLIC ChildCount : UINT //! Registered population starting at ChildArrayLowerBound; zero when unavailable.
GET // PUBLIC
ChildCount := 0;
IF NOT (FInitialized OR FCheckingInitialization) OR NOT FCollectionConfiguration.IsValid THEN
    RETURN;
END_IF;
ChildCount := FCollectionConfiguration.Count;
END_GET
END_PROPERTY

{region 'Documentation'}
(*!
<summary>Initializes and registers this owner's static Test Cases.</summary>
<description>
The owner identity is already established. Initialize owned children, bind the local interface
array through Builder.Initialize, select the mode, and use Register or RegisterWithSlot as
appropriate.

The base calls Finalize after this hook and retains only validated configuration values; it
then initializes the Orchestrator and calls CheckInitialization. Do not retain the borrowed
TestSuiteConfigurationBuilder or its temporary storage binding.

Implement GetTestCase against that same array and keep the composition fixed until full
hierarchical reinitialization. This abstract hook has no base implementation to call.
</description>
*)
{endregion}
METHOD PROTECTED ABSTRACT Configure
VAR_IN_OUT
    // SA0167: Borrowed builder; VAR_IN_OUT creates no temporary instance.
    {attribute 'analysis' := '-167'}
    Builder : TestSuiteConfigurationBuilder; //! Borrowed setup builder; initialize and register children during Configure only. The base calls Finalize afterwards.
END_VAR
(* Builder.Initialize(Mode := E_OrchestrationMode.Serial,
    TestCases := FTestCases);
FExample.Initialize(Parent := THIS^,
    TestName := 'Example',
    Config := ExampleConfig);
Builder.Register(TestCase := FExample);
Initialize and register each owned child. Use RegisterWithSlot for ParallelSlots.
The base calls Finalize after this method returns, including an early return.
Do not retain the builder or mutate the array after configuration.
*)
END_METHOD

{region 'Documentation'}
(*!
<summary>Publishes Result then Aggregation in the single Completing cycle, after result/status projection.</summary>
<description>
The single-call Completing phase provides one-shot Result then Aggregation publication; the next sequencing call enters Completed. Failed insertion is accounted for by the publisher without a retry here. Later child status changes do not rewrite the published payload.
</description>
*)
{endregion}
METHOD PRIVATE EmitFinalizationEvents
IF FState <> E_State.Completing THEN
    RETURN;
END_IF;

PublishEvent(Event := CreateResultEvent(OwnerScope := E_OwnerScope.TestSuite,
    Name := FName,
    ResourceName := FResourceName,
    State := FState,
    Result := FResult,
    Message := ''));
PublishEvent(Event := CreateTestSuiteAggregationEvent(Name := FName,
    ResourceName := FResourceName,
    Status := FStatus));
END_METHOD

{region 'Documentation'}
(*!
<summary>Latches the technical Suite error and emits its first diagnostic; does not change state.</summary>
*)
{endregion}
METHOD PRIVATE Error
VAR_INPUT
    Message : STRING(GVL_Constants.MessageLength); //! Framework diagnostic text emitted only when first escalating a mutable owner result to Error.
END_VAR
IF (FState = E_State.Uninitialized) OR (FState = E_State.Completed) THEN
    RETURN;
END_IF;
IF FResult <> E_Result.Error THEN
    PublishEvent(Event := CreateFrameworkEvent(Name := FName,
        ResourceName := FResourceName,
        State := FState,
        Severity := E_EventSeverity.Error,
        Message := Message));
END_IF;
FResult := E_Result.Error;
END_METHOD

{region 'Documentation'}
(*!
<summary>Returns this instance's retained event-publication service.</summary>
<description>
If the local binding is zero, the getter takes GVL_EventBuffer.Publisher on access. An
established binding is retained; Initialize and lifecycle Reset do not replace it.

The default must be bound before first diagnostic use. Controlled test adapters may assign the
protected field before use. This getter performs no event publication, lifecycle processing or
reservation change.
</description>
*)
{endregion}
{attribute 'monitoring' := 'variable'}
PROPERTY PUBLIC EventPublisher : I_EventPublisher //! Returns this instance's retained event-publication service.
GET // PUBLIC
IF FEventPublisher = 0 THEN
    FEventPublisher := GVL_EventBuffer.Publisher;
END_IF;
EventPublisher := FEventPublisher;
END_GET
END_PROPERTY

{region 'Documentation'}
(*!
<summary>Parent-assigned configuration slot; Initialize and Reset retain it.</summary>
*)
{endregion}
{attribute 'monitoring' := 'call'}
PROPERTY PUBLIC ExecutionSlot : UINT //! Parent-assigned configuration slot; Initialize and Reset retain it.
GET // PUBLIC
ExecutionSlot := FExecutionSlot;
END_GET
SET // PUBLIC
FExecutionSlot := ExecutionSlot;
END_SET
END_PROPERTY

